// Разрешения считаются только владельцем механизма.
Status.xConfirmAllowed := xRecovery
	AND Input.xPowered
	AND (uiCandidate <> UINT#0)
	AND (Error.dwErrorActive = DWORD#0);
Status.xStartAllowed := Status.xConfirmAllowed
	AND xRobotMagazineReady
	AND xPointsConfigured;
// Общая технологическая готовность не зависит от heartbeat HMI.
xEnableBaseAllowed := xBase
	AND xIdle
	AND Status.xConfirmed
	AND xRobotMagazineReady
	AND xPointsConfigured
	AND (uiCandidate = Status.uiRobotPallet)
	AND Input.xPowered
	AND (Error.dwErrorActive = DWORD#0);
Status.xEnableAllowed := xEnableBaseAllowed AND xConnection;
// Обмен не требует глобальной остановки робота: проверяется только отсутствие
// текущей или уже выданной операции именно с этим магазином.
Status.xSwapAllowed := xBase
	AND xConnection
	AND xIdle
	AND Input.xStandstill
	AND Input.xPowered
	AND (Error.dwErrorActive = DWORD#0)
	AND Status.xConfirmed
	AND (uiCandidate = Status.uiRobotPallet)
	AND NOT Status.xEnabled
	AND NOT xStopRequest
	AND xRobotSwapWindow;
xAutoSwapAllowed := xEnableBaseAllowed
	AND xRobotSwapWindow
	AND Status.xEnabled
	AND xOtherLoaded;
Status.xPowerAllowed := xRecovery
	AND NOT Input.xDriveError
	AND NOT xContradiction;
Status.xDriveResetAllowed := xSelected
	AND xManual
	AND xConnection
	AND Input.xAxisBound
	AND Input.xStandstill
	AND xIdle;
Status.xLowerAllowed := xPneumaticRecovery;
Status.xRaiseAllowed := xRecovery
	AND NOT xContradiction
	AND NOT Status.xHomeRequired;
Status.xSelectAllowed := xRecovery
	AND NOT xContradiction
	AND Input.xLiftDown
	AND NOT Input.xLiftUp
	AND xExchange;
// Наладочные команды замка и фиксатора независимы от подъёма и координаты.
// Это позволяет вернуть герконы в согласованное состояние после остановки.
Status.xLockAllowed := xPneumaticRecovery;
Status.xStopAllowed := xPneumaticRecovery;
Status.xHomeAllowed := xRecovery
	AND Input.xPowered
	AND NOT Input.xDriveError
	AND Input.xLiftDown
	AND NOT Input.xLiftUp
	AND xPairValid
	AND NOT xContradiction;
Status.xMoveAllowed := Status.xHomeAllowed
	AND Input.xHomed
	AND NOT Status.xHomeRequired;
Status.xJogAllowed := Status.xHomeAllowed;
Status.xTeachOperatorAllowed := Status.xMoveAllowed
	AND Input.xLiftDown
	AND NOT Input.xLiftUp;
Status.xTeachWorkAllowed := Status.xTeachOperatorAllowed
	AND ((uiSelected = UINT#1) OR (uiSelected = UINT#2));
Status.xResetAllowed := xRecovery
	AND (Error.dwErrorActive <> DWORD#0)
	AND NOT xContradiction
	AND NOT Input.xDriveError
	AND NOT Status.xHomeRequired
	AND xPairValid
	AND (Input.xLiftDown XOR Input.xLiftUp);
Status.xConfigAllowed := xSelected
	AND xManual
	AND xIdle
	AND NOT Status.xEnabled
	AND (Input.xStandstill OR NOT Input.xAxisBound)
	AND NOT Input.xPowered
	AND NOT xRobotOperation;

// Командный интерфейс FB не зависит от транспортных номеров HMI 1..19.
xCommandPresent := Command.xEnable
	OR Command.xConfirm
	OR Command.xStart
	OR Command.xRejectStart
	OR Command.xDisable
	OR Command.xSwap
	OR Command.xPowerOn
	OR Command.xPowerOff
	OR Command.xDriveReset
	OR Command.xHome
	OR Command.xLower
	OR Command.xRaise
	OR Command.xSelectPallet
	OR Command.xLockIn
	OR Command.xLockOut
	OR Command.xStopIn
	OR Command.xStopOut
	OR Command.xMoveToExchange
	OR Command.xMoveToWork
	OR Command.xStop
	OR Command.xReset
	OR Command.xJogPositive
	OR Command.xJogNegative
	OR Command.xJogRelease
	OR Command.xTeachOperator
	OR Command.xTeachWork;
xAccepted := NOT xCommandPresent;

IF Command.xStart THEN
	IF Status.xStartAllowed
		AND (Command.udiRevision = Status.udiRevision)
		AND (Command.uiPallet = uiCandidate) THEN
		Status.uiRobotPallet := uiCandidate;
		uiConfirmedCandidate := uiCandidate;
		Status.xConfirmed := TRUE;
		Status.xEnabled := TRUE;
		Status.rP1 := 0.0;
		Status.rP2 := 0.0;
		IF uiCandidate = UINT#1 THEN
			Status.rP1 := 1.0;
		ELSE
			Status.rP2 := 1.0;
		END_IF;
		xAccepted := TRUE;
	END_IF;
ELSIF Command.xRejectStart THEN
	Diag.stWarning.uiCode := WRN_START_REJECTED_BY_OPERATOR;
	Diag.stWarning.udiSequence := Diag.stWarning.udiSequence + UDINT#1;
	IF Diag.stWarning.udiSequence = UDINT#0 THEN
		Diag.stWarning.udiSequence := UDINT#1;
	END_IF;
	xAccepted := TRUE;
ELSIF Command.xEnable THEN
	IF Status.xEnableAllowed THEN
		Status.xEnabled := TRUE;
		xAccepted := TRUE;
	END_IF;
ELSIF Command.xConfirm THEN
	IF Status.xConfirmAllowed
		AND (Command.udiRevision = Status.udiRevision)
		AND (Command.uiPallet = uiCandidate) THEN
		Status.uiRobotPallet := uiCandidate;
		uiConfirmedCandidate := uiCandidate;
		Status.xConfirmed := TRUE;
		Status.rP1 := 0.0;
		Status.rP2 := 0.0;
		IF uiCandidate = UINT#1 THEN
			Status.rP1 := 1.0;
		ELSE
			Status.rP2 := 1.0;
		END_IF;
		xAccepted := TRUE;
	END_IF;
ELSIF Command.xDisable THEN
	Status.xEnabled := FALSE;
	xAccepted := TRUE;
ELSIF Command.xSwap THEN
	IF Status.xSwapAllowed THEN
		xExchangeStartedManual := xManual;
		Diag.eState := E_TWO_PALLET_STATE.AUTO_LOWER;
		xAccepted := TRUE;
	END_IF;
ELSIF Command.xPowerOn THEN
	IF Status.xPowerAllowed THEN
		Output.xPowerOn := TRUE;
		xAccepted := TRUE;
	END_IF;
ELSIF Command.xPowerOff THEN
	IF Status.xDriveResetAllowed THEN
		Output.xPowerOff := TRUE;
		Status.xConfirmed := FALSE;
		Status.xEnabled := FALSE;
		xAccepted := TRUE;
	END_IF;
ELSIF Command.xDriveReset THEN
	IF Status.xDriveResetAllowed AND Input.xDriveError THEN
		Output.xDriveReset := TRUE;
		Status.xConfirmed := FALSE;
		Status.xEnabled := FALSE;
		Status.xHomeRequired := TRUE;
		xAccepted := TRUE;
	END_IF;
ELSIF Command.xHome THEN
	IF Status.xHomeAllowed THEN
		Diag.eState := E_TWO_PALLET_STATE.MANUAL_HOME;
		xAccepted := TRUE;
	END_IF;
ELSIF Command.xLower THEN
	IF Status.xLowerAllowed THEN
		Diag.eState := E_TWO_PALLET_STATE.MANUAL_LOWER;
		xAccepted := TRUE;
	END_IF;
ELSIF Command.xRaise THEN
	IF Status.xRaiseAllowed THEN
		Diag.eState := E_TWO_PALLET_STATE.MANUAL_RAISE;
		xAccepted := TRUE;
	END_IF;
ELSIF Command.xSelectPallet THEN
	IF Status.xSelectAllowed
		AND ((Command.uiPallet = UINT#1) OR (Command.uiPallet = UINT#2)) THEN
		uiTo := Command.uiPallet;
		Diag.eState := E_TWO_PALLET_STATE.MANUAL_SELECT_PALLET;
		xAccepted := TRUE;
	END_IF;
ELSIF Command.xLockIn OR Command.xLockOut THEN
	IF Status.xLockAllowed THEN
		xManualLockOutTarget := Command.xLockOut;
		Diag.eState := E_TWO_PALLET_STATE.MANUAL_LOCK;
		xAccepted := TRUE;
	END_IF;
ELSIF Command.xStopIn OR Command.xStopOut THEN
	IF Status.xStopAllowed THEN
		xManualStopOutTarget := Command.xStopOut;
		Diag.eState := E_TWO_PALLET_STATE.MANUAL_STOP;
		xAccepted := TRUE;
	END_IF;
ELSIF Command.xMoveToExchange OR Command.xMoveToWork THEN
	IF Status.xMoveAllowed THEN
		lrTarget := Config.lrExchange;
		IF Command.xMoveToWork THEN
			lrTarget := lrWork;
		END_IF;
		Diag.eState := E_TWO_PALLET_STATE.MANUAL_MOVE;
		xAccepted := TRUE;
	END_IF;
ELSIF Command.xStop THEN
	Status.xEnabled := FALSE;
	// Stop неподвижного механизма не является ручным вмешательством.
	IF (Diag.eState <> E_TWO_PALLET_STATE.IDLE) OR (Input.xPowered AND NOT Input.xStandstill) THEN
		Output.xStop := TRUE;
		Status.xConfirmed := FALSE;
		Error.dwErrorActive := Error.dwErrorActive OR ERR_SEQUENCE_INTERRUPTED;
	END_IF;
	Diag.eState := E_TWO_PALLET_STATE.IDLE;
	uiJogDirection := UINT#0;
	xAccepted := TRUE;
ELSIF Command.xReset THEN
	IF Status.xResetAllowed THEN
		Error.dwErrorLast := Error.dwErrorActive;
		Error.dwErrorActive := DWORD#0;
		Status.xConfirmed := FALSE;
		Status.xEnabled := FALSE;
		xAccepted := TRUE;
	END_IF;
ELSIF Command.xJogPositive OR Command.xJogNegative THEN
	IF Status.xJogAllowed
		OR ((Diag.eState = E_TWO_PALLET_STATE.MANUAL_JOG)
			AND xBase
			AND xManual
			AND xConnection) THEN
		Diag.eState := E_TWO_PALLET_STATE.MANUAL_JOG;
		IF Command.xJogPositive THEN
			uiJogDirection := JOG_POSITIVE;
		ELSE
			uiJogDirection := JOG_NEGATIVE;
		END_IF;
		xAccepted := TRUE;
	END_IF;
ELSIF Command.xJogRelease THEN
	uiJogDirection := UINT#0;
	IF Diag.eState = E_TWO_PALLET_STATE.MANUAL_JOG THEN
		Diag.eState := E_TWO_PALLET_STATE.IDLE;
		Output.xStop := TRUE;
	END_IF;
	xAccepted := TRUE;
ELSIF Command.xTeachOperator THEN
	IF Status.xTeachOperatorAllowed THEN
		Output.xTeachOperator := TRUE;
		xAccepted := TRUE;
	END_IF;
ELSIF Command.xTeachWork THEN
	IF Status.xTeachWorkAllowed THEN
		Output.xTeachWork := TRUE;
		xAccepted := TRUE;
	END_IF;
END_IF;

IF xCommandPresent AND NOT xAccepted THEN
	IF (Command.xEnable OR Command.xStart) AND NOT xPointsConfigured THEN
		Diag.stWarning.uiCode := WRN_ENABLE_POINTS;
	ELSE
		Diag.stWarning.uiCode := WRN_COMMAND_REJECTED;
	END_IF;
	Diag.stWarning.udiSequence := Diag.stWarning.udiSequence + UDINT#1;
	IF Diag.stWarning.udiSequence = UDINT#0 THEN
		Diag.stWarning.udiSequence := UDINT#1;
	END_IF;
END_IF;

IF xExternalCommandRejected THEN
	Diag.stWarning.uiCode := WRN_COMMAND_REJECTED;
	Diag.stWarning.udiSequence := Diag.stWarning.udiSequence + UDINT#1;
	IF Diag.stWarning.udiSequence = UDINT#0 THEN
		Diag.stWarning.udiSequence := UDINT#1;
	END_IF;
END_IF;

Status.xCommandAccepted := xAccepted;

IF xAutoSwap
	AND xAutoSwapAllowed
	AND NOT Output.xStop
	AND NOT xCommandPresent THEN
	xExchangeStartedManual := FALSE;
	Diag.eState := E_TWO_PALLET_STATE.AUTO_LOWER;
END_IF;

// Стоп ячейки имеет приоритет над командой, принятой в том же скане.
// В IDLE при остановленной оси сохраняем включение и подтверждение.
// Собственные Command.xStop / Command.xDisable отдельно отключают магазин.
IF xStopRequest THEN
	IF (Diag.eState <> E_TWO_PALLET_STATE.IDLE) OR (Input.xPowered AND NOT Input.xStandstill) THEN
		Error.dwErrorActive := Error.dwErrorActive OR ERR_SEQUENCE_INTERRUPTED;
		Output.xStop := TRUE;
		Status.xConfirmed := FALSE;
		Status.xEnabled := FALSE;
	END_IF;
	Diag.eState := E_TWO_PALLET_STATE.IDLE;
END_IF;

// Команда могла сменить состояние в этом же скане — обновляем классификацию
// до обработки входа в шаг и запуска таймеров.
xAutomaticState := (Diag.eState = E_TWO_PALLET_STATE.AUTO_LOWER)
	OR (Diag.eState = E_TWO_PALLET_STATE.AUTO_MOVE_TO_EXCHANGE)
	OR (Diag.eState = E_TWO_PALLET_STATE.AUTO_SELECT_PALLET)
	OR (Diag.eState = E_TWO_PALLET_STATE.AUTO_MOVE_TO_WORK)
	OR (Diag.eState = E_TWO_PALLET_STATE.AUTO_RAISE);
xManualState := (Diag.eState = E_TWO_PALLET_STATE.MANUAL_LOWER)
	OR (Diag.eState = E_TWO_PALLET_STATE.MANUAL_RAISE)
	OR (Diag.eState = E_TWO_PALLET_STATE.MANUAL_SELECT_PALLET)
	OR (Diag.eState = E_TWO_PALLET_STATE.MANUAL_MOVE)
	OR (Diag.eState = E_TWO_PALLET_STATE.MANUAL_HOME)
	OR (Diag.eState = E_TWO_PALLET_STATE.MANUAL_JOG)
	OR (Diag.eState = E_TWO_PALLET_STATE.MANUAL_LOCK)
	OR (Diag.eState = E_TWO_PALLET_STATE.MANUAL_STOP);
xManualPneumaticState := (Diag.eState = E_TWO_PALLET_STATE.MANUAL_LOWER)
	OR (Diag.eState = E_TWO_PALLET_STATE.MANUAL_LOCK)
	OR (Diag.eState = E_TWO_PALLET_STATE.MANUAL_STOP);

IF (Diag.eState = E_TWO_PALLET_STATE.AUTO_LOWER)
	AND (ePreviousState <> E_TWO_PALLET_STATE.AUTO_LOWER) THEN
	uiFrom := Status.uiRobotPallet;
	uiTo := UINT#3 - uiFrom;
END_IF;

xStateEntry := Diag.eState <> ePreviousState;
IF xManualState AND xStateEntry THEN
	Status.xConfirmed := FALSE;
	Status.xEnabled := FALSE;
	Status.udiRevision := Status.udiRevision + UDINT#1;
	IF Status.udiRevision = UDINT#0 THEN
		Status.udiRevision := UDINT#1;
	END_IF;
END_IF;

IF xStateEntry THEN
	xSeenMotion := FALSE;
	xSeenDone := FALSE;
	IF (Diag.eState = E_TWO_PALLET_STATE.MANUAL_MOVE)
		OR (Diag.eState = E_TWO_PALLET_STATE.MANUAL_HOME)
		OR (Diag.eState = E_TWO_PALLET_STATE.MANUAL_JOG) THEN
		uiManualSelected := uiSelected;
	END_IF;
ELSIF Input.xMotionDone THEN
	xSeenDone := TRUE;
END_IF;

IF NOT Input.xStandstill THEN
	xSeenMotion := TRUE;
END_IF;

tStateLimit := Config.tCylinder;
IF (Diag.eState = E_TWO_PALLET_STATE.AUTO_MOVE_TO_EXCHANGE)
	OR (Diag.eState = E_TWO_PALLET_STATE.AUTO_MOVE_TO_WORK)
	OR (Diag.eState = E_TWO_PALLET_STATE.MANUAL_MOVE) THEN
	tStateLimit := Config.tMove;
END_IF;
IF Diag.eState = E_TWO_PALLET_STATE.MANUAL_HOME THEN
	tStateLimit := Config.tHome;
END_IF;

tonState(
	IN := NOT xIdle
		AND (Diag.eState <> E_TWO_PALLET_STATE.MANUAL_JOG)
		AND NOT xStateEntry,
	PT := tStateLimit);
tonCoil(
	IN := NOT xIdle AND NOT xStateEntry,
	PT := Config.tPulse);
tonJogLease(
	IN := (Diag.eState = E_TWO_PALLET_STATE.MANUAL_JOG)
		AND NOT (Command.xJogPositive OR Command.xJogNegative),
	PT := T#350MS);
ePreviousState := Diag.eState;

// Автомат обмена и ручного восстановления.
uiTargetSignals := Config.uiP1Signals;
IF uiTo = UINT#2 THEN uiTargetSignals := Config.uiP2Signals; END_IF;
CASE Diag.eState OF
	E_TWO_PALLET_STATE.AUTO_LOWER,
	E_TWO_PALLET_STATE.MANUAL_LOWER:
		xLiftDownCommand := TRUE;
		IF Input.xLiftDown AND NOT Input.xLiftUp THEN
			IF Diag.eState = E_TWO_PALLET_STATE.AUTO_LOWER THEN
				Diag.eState := E_TWO_PALLET_STATE.AUTO_MOVE_TO_EXCHANGE;
				lrTarget := Config.lrExchange;
			ELSE
				Diag.eState := E_TWO_PALLET_STATE.IDLE;
			END_IF;
		END_IF;

	E_TWO_PALLET_STATE.AUTO_MOVE_TO_EXCHANGE,
	E_TWO_PALLET_STATE.AUTO_MOVE_TO_WORK,
	E_TWO_PALLET_STATE.MANUAL_MOVE:
		IF Diag.eState = E_TWO_PALLET_STATE.AUTO_MOVE_TO_WORK THEN
			lrTarget := Config.lrWorkP1;
			IF uiTo = UINT#2 THEN
				lrTarget := Config.lrWorkP2;
			END_IF;
		END_IF;

		IF NOT Input.xLiftDown
			OR Input.xLiftUp
			OR NOT xPairValid
			OR Status.xHomeRequired
			OR ((Diag.eState = E_TWO_PALLET_STATE.AUTO_MOVE_TO_EXCHANGE) AND (uiSelected <> uiFrom))
			OR ((Diag.eState = E_TWO_PALLET_STATE.AUTO_MOVE_TO_WORK) AND (uiSelected <> uiTo))
			OR ((Diag.eState = E_TWO_PALLET_STATE.MANUAL_MOVE) AND (uiSelected <> uiManualSelected))
			OR (Input.xLimitPositive AND (lrTarget > Input.lrPosition + Config.lrTolerance))
			OR (Input.xLimitNegative AND (lrTarget < Input.lrPosition - Config.lrTolerance)) THEN
			Error.dwErrorActive := Error.dwErrorActive OR ERR_LOGIC;
			Diag.eState := E_TWO_PALLET_STATE.IDLE;
			Output.xStop := TRUE;
		ELSE
			Output.lrTarget := lrTarget;
			Output.xMove := xStateEntry;
			IF Input.xStandstill
				AND (ABS(Input.lrPosition - lrTarget) <= Config.lrTolerance)
				AND ((xSeenMotion OR xSeenDone) OR xStateEntry) THEN
				Output.xMove := FALSE;
				IF Diag.eState = E_TWO_PALLET_STATE.AUTO_MOVE_TO_EXCHANGE THEN
					Diag.eState := E_TWO_PALLET_STATE.AUTO_SELECT_PALLET;
				ELSIF Diag.eState = E_TWO_PALLET_STATE.AUTO_MOVE_TO_WORK THEN
					Diag.eState := E_TWO_PALLET_STATE.AUTO_RAISE;
				ELSE
					Diag.eState := E_TWO_PALLET_STATE.IDLE;
				END_IF;
			END_IF;
		END_IF;

	E_TWO_PALLET_STATE.AUTO_SELECT_PALLET,
	E_TWO_PALLET_STATE.MANUAL_SELECT_PALLET:
		IF NOT xExchange OR NOT Input.xLiftDown OR Input.xLiftUp THEN
			Error.dwErrorActive := Error.dwErrorActive OR ERR_LOGIC;
			Diag.eState := E_TWO_PALLET_STATE.IDLE;
			Output.xStop := TRUE;
		ELSE
			xSelectCommand := TRUE;
		END_IF;
		IF (uiSelected = uiTo) AND xPairValid AND NOT Output.xStop THEN
			IF Diag.eState = E_TWO_PALLET_STATE.AUTO_SELECT_PALLET THEN
				Diag.eState := E_TWO_PALLET_STATE.AUTO_MOVE_TO_WORK;
			ELSE
				Diag.eState := E_TWO_PALLET_STATE.IDLE;
			END_IF;
		END_IF;

	E_TWO_PALLET_STATE.MANUAL_LOCK:
		IF xManualLockOutTarget THEN
			xManualLockCommand := NOT Input.xLockOut OR Input.xLockIn;
			IF Input.xLockOut AND NOT Input.xLockIn THEN Diag.eState := E_TWO_PALLET_STATE.IDLE; END_IF;
		ELSE
			xManualLockCommand := NOT Input.xLockIn OR Input.xLockOut;
			IF Input.xLockIn AND NOT Input.xLockOut THEN Diag.eState := E_TWO_PALLET_STATE.IDLE; END_IF;
		END_IF;

	E_TWO_PALLET_STATE.MANUAL_STOP:
		IF xManualStopOutTarget THEN
			xManualStopCommand := NOT Input.xStopOut OR Input.xStopIn;
			IF Input.xStopOut AND NOT Input.xStopIn THEN Diag.eState := E_TWO_PALLET_STATE.IDLE; END_IF;
		ELSE
			xManualStopCommand := NOT Input.xStopIn OR Input.xStopOut;
			IF Input.xStopIn AND NOT Input.xStopOut THEN Diag.eState := E_TWO_PALLET_STATE.IDLE; END_IF;
		END_IF;

	E_TWO_PALLET_STATE.AUTO_RAISE:
		// Завершение обмена устанавливает подъём по выбранной конфигурации
		// только после фактического останова в рабочей позиции.
		IF NOT xWork
			OR Status.xHomeRequired
			OR (uiSelected <> uiTo) THEN
			Error.dwErrorActive := Error.dwErrorActive OR ERR_LOGIC;
			Diag.eState := E_TWO_PALLET_STATE.IDLE;
			Output.xStop := TRUE;
		ELSE
			xLiftUpCommand := (uiTargetSignals AND UINT#2) <> UINT#0;
			xLiftDownCommand := NOT xLiftUpCommand;
			IF uiSignals = uiTargetSignals THEN
				Status.uiRobotPallet := uiTo;
				uiConfirmedCandidate := uiTo;
				Status.xConfirmed := TRUE;
				Status.xCompleted := TRUE;
				Diag.eState := E_TWO_PALLET_STATE.IDLE;
			END_IF;
		END_IF;

	E_TWO_PALLET_STATE.MANUAL_RAISE:
		// Наладочный подъём не требует HOME-координаты или рабочей позиции.
		IF NOT Input.xStandstill OR NOT xManual OR xContradiction OR Status.xHomeRequired THEN
			Error.dwErrorActive := Error.dwErrorActive OR ERR_LOGIC;
			Diag.eState := E_TWO_PALLET_STATE.IDLE;
			Output.xStop := TRUE;
		ELSE
			xLiftUpCommand := TRUE;
			IF Input.xLiftUp AND NOT Input.xLiftDown THEN
				Diag.eState := E_TWO_PALLET_STATE.IDLE;
			END_IF;
		END_IF;

	E_TWO_PALLET_STATE.MANUAL_HOME:
		Output.xHome := xStateEntry;
		IF xSeenDone
			AND Input.xHomed
			AND Input.xStandstill
			AND NOT xStateEntry THEN
			Status.xHomeRequired := FALSE;
			Diag.eState := E_TWO_PALLET_STATE.IDLE;
		END_IF;

	E_TWO_PALLET_STATE.MANUAL_JOG:
		IF tonJogLease.Q OR NOT xConnection OR (uiJogDirection = UINT#0) THEN
			Diag.eState := E_TWO_PALLET_STATE.IDLE;
			Output.xStop := TRUE;
		ELSE
			Output.xJogPositive := (uiJogDirection = JOG_POSITIVE) AND NOT Input.xLimitPositive;
			Output.xJogNegative := (uiJogDirection = JOG_NEGATIVE) AND NOT Input.xLimitNegative;
		END_IF;

	E_TWO_PALLET_STATE.IDLE:
		uiJogDirection := UINT#0;

ELSE
	Error.dwErrorActive := Error.dwErrorActive OR ERR_LOGIC;
	Diag.eState := E_TWO_PALLET_STATE.IDLE;
	Output.xStop := TRUE;
END_CASE;
IF Diag.eState = E_TWO_PALLET_STATE.IDLE THEN xExchangeStartedManual := FALSE; END_IF;

// Низ П2 и выбранное зацепление контролируются всё время Home/JOG.
IF ((Diag.eState = E_TWO_PALLET_STATE.MANUAL_HOME)
	OR (Diag.eState = E_TWO_PALLET_STATE.MANUAL_JOG))
	AND (NOT Input.xLiftDown
		OR Input.xLiftUp
		OR NOT xPairValid
		OR (uiSelected <> uiManualSelected)
		OR xContradiction
		OR Input.xDriveError
		OR NOT Input.xPowered) THEN
	Error.dwErrorActive := Error.dwErrorActive OR ERR_LOGIC;
	Diag.eState := E_TWO_PALLET_STATE.IDLE;
	Output.xStop := TRUE;
END_IF;

IF tonState.Q THEN
	IF (ePreviousState = E_TWO_PALLET_STATE.AUTO_MOVE_TO_EXCHANGE)
		OR (ePreviousState = E_TWO_PALLET_STATE.AUTO_MOVE_TO_WORK)
		OR (ePreviousState = E_TWO_PALLET_STATE.MANUAL_MOVE)
		OR (ePreviousState = E_TWO_PALLET_STATE.MANUAL_HOME) THEN
		Error.dwErrorActive := Error.dwErrorActive OR ERR_MOTION_TIMEOUT;
		Status.xHomeRequired := TRUE;
	ELSE
		Error.dwErrorActive := Error.dwErrorActive OR ERR_CYLINDER_TIMEOUT;
	END_IF;
	Diag.eState := E_TWO_PALLET_STATE.IDLE;
	Output.xStop := TRUE;
END_IF;

IF (((NOT xBase) AND NOT (xManualPneumaticState AND xPneumaticBase))
	OR ((NOT xConnection) AND xManualState AND NOT xManualPneumaticState))
	AND (ePreviousState <> E_TWO_PALLET_STATE.IDLE)
	OR Output.xStop THEN
	Output.xMove := FALSE;
	Output.xHome := FALSE;
	Output.xJogPositive := FALSE;
	Output.xJogNegative := FALSE;
	xLiftUpCommand := FALSE;
	xLiftDownCommand := FALSE;
	xSelectCommand := FALSE;
	xManualLockCommand := FALSE;
	xManualStopCommand := FALSE;
END_IF;

// Автоматический обмен переключает пару совместно; ручное восстановление — каждый цилиндр отдельно.
xLockOutTarget := (uiTargetSignals AND UINT#8) <> UINT#0;
xStopOutTarget := (uiTargetSignals AND UINT#32) <> UINT#0;
Output.xLiftUp := xBase AND xLiftUpCommand AND NOT tonCoil.Q;
Output.xLiftDown := (xBase OR xPneumaticBase) AND xLiftDownCommand AND NOT tonCoil.Q;
Output.xLockOut := (xBase AND xSelectCommand AND xLockOutTarget
	OR xPneumaticBase AND xManualLockCommand AND xManualLockOutTarget) AND NOT tonCoil.Q;
Output.xLockIn := (xBase AND xSelectCommand AND NOT xLockOutTarget
	OR xPneumaticBase AND xManualLockCommand AND NOT xManualLockOutTarget) AND NOT tonCoil.Q;
Output.xStopOut := (xBase AND xSelectCommand AND xStopOutTarget
	OR xPneumaticBase AND xManualStopCommand AND xManualStopOutTarget) AND NOT tonCoil.Q;
Output.xStopIn := (xBase AND xSelectCommand AND NOT xStopOutTarget
	OR xPneumaticBase AND xManualStopCommand AND NOT xManualStopOutTarget) AND NOT tonCoil.Q;

// Поза для 3D — оценка по координате каретки и подтверждённому зацеплению.
IF xPairValid AND Input.xHomed THEN
	lrSpan := lrWork - Config.lrExchange;
	IF ABS(lrSpan) > Config.lrTolerance THEN
		rTravel := LREAL_TO_REAL(
			LIMIT(0.0, (Input.lrPosition - Config.lrExchange) / lrSpan, 1.0));
		IF uiSelected = UINT#1 THEN
			Status.rP1 := rTravel;
		ELSE
			Status.rP2 := rTravel;
		END_IF;
	END_IF;
END_IF;

IF Input.xLiftUp AND NOT Input.xLiftDown THEN
	Status.rLift := 1.0;
ELSIF Input.xLiftDown AND NOT Input.xLiftUp THEN
	Status.rLift := 0.0;
END_IF;

// Диагностика и совместимый публичный Status формируются в одном месте.
IF (Error.dwErrorActive <> dwPreviousError)
	AND (Error.dwErrorActive <> DWORD#0) THEN
	Diag.eFaultState := ePreviousState;
END_IF;
dwPreviousError := Error.dwErrorActive;

IF Error.dwErrorActive <> DWORD#0 THEN
	Error.dwErrorLast := Error.dwErrorActive;
	Status.xConfirmed := FALSE;
	Status.xEnabled := FALSE;
END_IF;
Error.dwAlarmActive := Error.dwErrorActive;
Error.stErrorActive := UpdateErrorView(dwError := Error.dwErrorActive);
Error.stErrorLast := UpdateErrorView(dwError := Error.dwErrorLast);

Status.uiStep := TO_UINT(Diag.eState);
Status.uiFaultStep := TO_UINT(Diag.eFaultState);
Status.uiReason := Diag.uiReason;
Status.dwError := Error.dwErrorActive;
Status.stWarning := Diag.stWarning;
Status.xBusy := Diag.eState <> E_TWO_PALLET_STATE.IDLE;
Status.xError := Error.dwErrorActive <> DWORD#0;

// Команда или автомат могли занять механизм после первоначального расчёта
// разрешений. Не публикуем устаревшее разрешение ещё на один скан.
IF Status.xBusy THEN
	Status.xConfirmAllowed := FALSE;
	Status.xStartAllowed := FALSE;
	Status.xEnableAllowed := FALSE;
	Status.xSwapAllowed := FALSE;
	Status.xPowerAllowed := FALSE;
	Status.xDriveResetAllowed := FALSE;
	Status.xHomeAllowed := FALSE;
	Status.xLowerAllowed := FALSE;
	Status.xRaiseAllowed := FALSE;
	Status.xSelectAllowed := FALSE;
	Status.xLockAllowed := FALSE;
	Status.xStopAllowed := FALSE;
	Status.xMoveAllowed := FALSE;
	Status.xJogAllowed := FALSE;
	Status.xTeachOperatorAllowed := FALSE;
	Status.xTeachWorkAllowed := FALSE;
	Status.xResetAllowed := FALSE;
	Status.xConfigAllowed := FALSE;
END_IF;

// Инвентарь операторской палеты редактируется всегда, независимо от режима,
// движения, подтверждения, питания и ошибок механизма. Роботная палета — только
// при выключенном магазине после освобождения текущей/выданной операции с ним.
// Считаем после команд и обмена, чтобы роль палеты была актуальна в этом скане.
Status.xEdit1Allowed := xSelected
	AND ((Status.uiRobotPallet <> UINT#1) OR (NOT Status.xEnabled AND xActivePalletEditAllowed));
Status.xEdit2Allowed := xSelected
	AND ((Status.uiRobotPallet <> UINT#2) OR (NOT Status.xEnabled AND xActivePalletEditAllowed));
Status.xEditAllowed := Status.xEdit1Allowed OR Status.xEdit2Allowed;
Status.xLoadAllowed := Status.xConfirmed AND NOT Status.xBusy AND NOT xOtherLoaded
	AND (((Status.uiRobotPallet = UINT#1) AND Status.xEdit2Allowed)
		OR ((Status.uiRobotPallet = UINT#2) AND Status.xEdit1Allowed));

Status.xReady := xSelected
	AND Status.xEnabled
	AND Status.xConfirmed
	AND NOT Status.xBusy
	AND NOT Status.xError
	AND xWork
	AND (uiCandidate = Status.uiRobotPallet)
	AND Input.xPowered
	AND xRobotGeometryReady
	AND xRobotMagazineReady
	AND xSafe;

IF NOT xSelected THEN
	Status.xEnabled := FALSE;
	Status.xConfirmed := FALSE;
END_IF;

METHOD IsSignalConfigurationValid : BOOL
VAR_INPUT
	uiP1Signals : UINT;
	uiP2Signals : UINT;
END_VAR
// Рабочее положение каждого цилиндра подтверждает ровно один геркон.
// Зацепление должно различать палеты и при опущенной П2 во время обмена.
IsSignalConfigurationValid := (uiP1Signals <= UINT#63)
	AND (uiP2Signals <= UINT#63)
	AND (((uiP1Signals AND UINT#3) = UINT#1) OR ((uiP1Signals AND UINT#3) = UINT#2))
	AND (((uiP2Signals AND UINT#3) = UINT#1) OR ((uiP2Signals AND UINT#3) = UINT#2))
	AND (((uiP1Signals AND UINT#12) = UINT#4) OR ((uiP1Signals AND UINT#12) = UINT#8))
	AND (((uiP2Signals AND UINT#12) = UINT#4) OR ((uiP2Signals AND UINT#12) = UINT#8))
	AND (((uiP1Signals AND UINT#48) = UINT#16) OR ((uiP1Signals AND UINT#48) = UINT#32))
	AND (((uiP2Signals AND UINT#48) = UINT#16) OR ((uiP2Signals AND UINT#48) = UINT#32))
	AND ((uiP1Signals AND UINT#60) <> (uiP2Signals AND UINT#60));
END_METHOD

METHOD UpdateErrorView : ST_TWO_PALLET_ERROR
VAR_INPUT
	dwError : DWORD;
END_VAR
VAR
	stError : ST_TWO_PALLET_ERROR;
END_VAR
stError.DRIVE_ERROR := (dwError AND ERR_DRIVE) <> DWORD#0;
stError.SENSOR_CONTRADICTION := (dwError AND ERR_SENSOR_CONTRADICTION) <> DWORD#0;
stError.CYLINDER_TIMEOUT := (dwError AND ERR_CYLINDER_TIMEOUT) <> DWORD#0;
stError.MOTION_TIMEOUT := (dwError AND ERR_MOTION_TIMEOUT) <> DWORD#0;
stError.LOGIC_ERROR := (dwError AND ERR_LOGIC) <> DWORD#0;
stError.SEQUENCE_INTERRUPTED := (dwError AND ERR_SEQUENCE_INTERRUPTED) <> DWORD#0;

UpdateErrorView := stError;
END_METHOD

END_FUNCTION_BLOCK

// Device/Application/FB/FB_TWO_PALLET_SIMULATION
FUNCTION_BLOCK FB_TWO_PALLET_SIMULATION
VAR_INPUT
	xEnable : BOOL; // Только тестовая среда SIMULATION
	uiP1Signals : UINT;
	Command : ST_TWO_PALLET_OUTPUT;
END_VAR
VAR_OUTPUT
	xLiftDown : BOOL;
	xLiftUp : BOOL;
	xLockIn : BOOL;
	xLockOut : BOOL;
	xStopIn : BOOL;
	xStopOut : BOOL;
END_VAR
VAR
	xInitialized : BOOL;
	xLiftTargetUp : BOOL;
	xLockTargetOut : BOOL;
	xStopTargetOut : BOOL;
	tonLift : TON;
	tonLock : TON;
	tonStop : TON;
END_VAR

IF NOT xEnable THEN
	xInitialized := FALSE;
	xLiftDown := FALSE;
	xLiftUp := FALSE;
	xLockIn := FALSE;
	xLockOut := FALSE;
	xStopIn := FALSE;
	xStopOut := FALSE;
	tonLift(IN := FALSE, PT := T#300MS);
	tonLock(IN := FALSE, PT := T#300MS);
	tonStop(IN := FALSE, PT := T#300MS);
ELSE
	IF NOT xInitialized THEN
		// Виртуальная начальная поза: П2 внизу, замок держит П1,
		// фиксатор держит противоположную палету.
		xLiftTargetUp := FALSE;
		xLockTargetOut := (uiP1Signals AND UINT#8) <> UINT#0;
		xStopTargetOut := (uiP1Signals AND UINT#32) <> UINT#0;
		xLiftDown := TRUE;
		xLiftUp := FALSE;
		xLockOut := xLockTargetOut;
		xLockIn := NOT xLockTargetOut;
		xStopOut := xStopTargetOut;
		xStopIn := NOT xStopTargetOut;
		xInitialized := TRUE;
	END_IF;

	// Бистабильный 5/2 сохраняет положение после снятия обеих катушек.
	IF Command.xLiftUp AND NOT Command.xLiftDown THEN
		xLiftTargetUp := TRUE;
	ELSIF Command.xLiftDown AND NOT Command.xLiftUp THEN
		xLiftTargetUp := FALSE;
	END_IF;
	IF Command.xLockOut AND NOT Command.xLockIn THEN
		xLockTargetOut := TRUE;
	ELSIF Command.xLockIn AND NOT Command.xLockOut THEN
		xLockTargetOut := FALSE;
	END_IF;
	IF Command.xStopOut AND NOT Command.xStopIn THEN
		xStopTargetOut := TRUE;
	ELSIF Command.xStopIn AND NOT Command.xStopOut THEN
		xStopTargetOut := FALSE;
	END_IF;

	tonLift(IN := xLiftTargetUp <> xLiftUp, PT := T#300MS);
	tonLock(IN := xLockTargetOut <> xLockOut, PT := T#300MS);
	tonStop(IN := xStopTargetOut <> xStopOut, PT := T#300MS);
	IF tonLift.Q THEN
		xLiftUp := xLiftTargetUp;
		xLiftDown := NOT xLiftTargetUp;
	END_IF;
	IF tonLock.Q THEN
		xLockOut := xLockTargetOut;
		xLockIn := NOT xLockTargetOut;
	END_IF;
	IF tonStop.Q THEN
		xStopOut := xStopTargetOut;
		xStopIn := NOT xStopTargetOut;
	END_IF;
END_IF;

END_FUNCTION_BLOCK

// Device/Application/FB/FB_MULTI_TYPE/FB_MULTI_TYPE_CONFIG_MANAGER
FUNCTION_BLOCK FB_MULTI_TYPE_CONFIG_MANAGER
VAR_INPUT
	xTestInitialize  : BOOL; // Атомарная загрузка конфигурации из тестового буфера
	stTestScenario   : ST_TEST_SCENARIO_BUFFER;
	Command          : ST_MULTI_TYPE_COMMAND; // Запросы конфигурации от HMI
	xCellRunning     : BOOL; // Автоматический цикл выполняется
	xMotionBusy      : BOOL; // Оси ещё движутся
	stRobotStatus    : ST_ROBOT_STATUS; // Состояние робота
	astMagazineStatus : ARRAY [1..GVL_CELL_SETTINGS.MagazineCount] OF ST_MAGAZINE_STATUS; // Оба магазина
	astMachineStatus : ARRAY [1..3] OF ST_MACHINE_PUBLIC; // Состояния станков
	uiRows           : UINT; // Строки активной матрицы
	uiColumns        : UINT; // Столбцы активной матрицы
END_VAR
VAR_OUTPUT
	Config : ST_MULTI_TYPE_CONFIG; // Фактически принятая конфигурация
	Status : ST_MULTI_TYPE_CONFIG_STATUS; // Разрешения и диагностика
END_VAR
VAR
	xInitialized        : BOOL; // Начальные безопасные значения заданы
	xAllMachinesSafe    : BOOL; // Станки не обслуживаются и не обрабатывают
	xAllMachinesDisabled: BOOL; // Все станки выключены
	xAllMagazinesEditable : BOOL; // Оба магазина выключены и не заняты
	xAllTypesHaveMachines : BOOL; // Каждый тип назначен хотя бы одному станку
	uiMachine           : UINT; // Индекс станка
	uiMagazine          : UINT; // Индекс магазина
	uiSlot              : UINT; // Индекс слота
	uiType              : UINT; // Индекс типа
	auiMachineCount     : ARRAY [1..3] OF UINT; // Количество станков каждого типа
	auiSlotCount        : ARRAY [1..3] OF UINT; // Количество слотов каждого типа
	rtSetTypeCount      : R_TRIG; // Фронт изменения количества типов
	rtSetMachineType    : R_TRIG; // Фронт назначения типа станку
	rtSetSlotType       : R_TRIG; // Фронт назначения типа слоту
	rtAutoDistribute    : R_TRIG; // Фронт автоматического распределения
END_VAR
VAR CONSTANT
	FIRST_MACHINE : UINT := UINT#1;
	LAST_MACHINE  : UINT := UINT#3;
	FIRST_TYPE    : UINT := UINT#1;
	LAST_TYPE     : UINT := UINT#3;
	WRN_TYPE_COUNT_NOT_ALLOWED : UINT := UINT#23;
	WRN_MACHINE_TYPE_REJECTED  : UINT := UINT#24;
	WRN_SLOT_TYPE_REJECTED     : UINT := UINT#25;
	WRN_DISTRIBUTION_REJECTED  : UINT := UINT#26;
END_VAR

IF (uiRows > UINT#0)
AND (uiColumns > UINT#0)
AND ((uiRows * uiColumns) <= SINT_TO_UINT(GVL_CELL_SETTINGS.NumberDetail)) THEN
	Status.uiActiveSlotCount := uiRows * uiColumns;
ELSE
	Status.uiActiveSlotCount := UINT#0;
END_IF;

IF NOT xInitialized THEN
	Config.uiTypeCount := UINT#1;
	FOR uiMachine := FIRST_MACHINE TO LAST_MACHINE DO
		Config.auiMachineType[uiMachine] := UINT#1;
	END_FOR;
	FOR uiSlot := UINT#1 TO SINT_TO_UINT(GVL_CELL_SETTINGS.NumberDetail) DO
		IF uiSlot <= Status.uiActiveSlotCount THEN
			Config.auiSlotType[uiSlot] := UINT#1;
		ELSE
			Config.auiSlotType[uiSlot] := UINT#0;
		END_IF;
	END_FOR;
	xInitialized := TRUE;
END_IF;

xAllMachinesSafe := TRUE;
xAllMachinesDisabled := TRUE;
FOR uiMachine := FIRST_MACHINE TO LAST_MACHINE DO
	IF astMachineStatus[uiMachine].xBusy
	OR astMachineStatus[uiMachine].xProcessing THEN
		xAllMachinesSafe := FALSE;
	END_IF;
	IF astMachineStatus[uiMachine].xEnabled
	OR astMachineStatus[uiMachine].xDisablePending THEN
		xAllMachinesDisabled := FALSE;
	END_IF;
END_FOR;

xAllMagazinesEditable := TRUE;
FOR uiMagazine := UINT#1 TO INT_TO_UINT(GVL_CELL_SETTINGS.MagazineCount) DO
	IF astMagazineStatus[uiMagazine].xEnabled
	OR astMagazineStatus[uiMagazine].xBusy
	OR astMagazineStatus[uiMagazine].xDisablePending THEN
		xAllMagazinesEditable := FALSE;
	END_IF;
END_FOR;

Status.xMagazineConfigAllowed := NOT xCellRunning
	AND NOT xMotionBusy
	AND NOT stRobotStatus.xBusy
	AND NOT stRobotStatus.xBlankAvailable
	AND NOT stRobotStatus.xDetailAvailable
	AND xAllMagazinesEditable
	AND xAllMachinesSafe;
Status.xTypeCountAllowed := Status.xMagazineConfigAllowed
	AND xAllMachinesDisabled;

FOR uiMachine := FIRST_MACHINE TO LAST_MACHINE DO
	Status.axMachineTypeAllowed[uiMachine] := NOT xCellRunning
		AND NOT xMotionBusy
		AND NOT stRobotStatus.xBusy
		AND NOT stRobotStatus.xBlankAvailable
		AND NOT stRobotStatus.xDetailAvailable
		AND xAllMagazinesEditable
		AND NOT astMachineStatus[uiMachine].xEnabled
		AND NOT astMachineStatus[uiMachine].xDisablePending
		AND NOT astMachineStatus[uiMachine].xBusy
		AND NOT astMachineStatus[uiMachine].xProcessing;
END_FOR;

rtSetTypeCount(CLK := Command.xSetTypeCount);
rtSetMachineType(CLK := Command.xSetMachineType);
rtSetSlotType(CLK := Command.xSetSlotType);
rtAutoDistribute(CLK := Command.xAutoDistribute);

IF rtSetTypeCount.Q THEN
	IF NOT Status.xTypeCountAllowed
	OR (Command.uiRequestedTypeCount < FIRST_TYPE)
	OR (Command.uiRequestedTypeCount > LAST_TYPE) THEN
		RaiseWarning(uiCode := WRN_TYPE_COUNT_NOT_ALLOWED);
	ELSE
		Config.uiTypeCount := Command.uiRequestedTypeCount;
		CASE Config.uiTypeCount OF
			UINT#1:
				Config.auiMachineType[1] := UINT#1;
				Config.auiMachineType[2] := UINT#1;
				Config.auiMachineType[3] := UINT#1;
			UINT#2:
				Config.auiMachineType[1] := UINT#1;
				Config.auiMachineType[2] := UINT#1;
				Config.auiMachineType[3] := UINT#2;
			UINT#3:
				Config.auiMachineType[1] := UINT#1;
				Config.auiMachineType[2] := UINT#2;
				Config.auiMachineType[3] := UINT#3;
		END_CASE;
		ApplyDistribution();
	END_IF;
END_IF;

IF rtSetMachineType.Q THEN
	IF (Command.uiRequestedMachine < FIRST_MACHINE)
	OR (Command.uiRequestedMachine > LAST_MACHINE) THEN
		RaiseWarning(uiCode := WRN_MACHINE_TYPE_REJECTED);
	ELSE
		IF (Command.uiRequestedMachineType < FIRST_TYPE)
		OR (Command.uiRequestedMachineType > Config.uiTypeCount)
		OR NOT Status.axMachineTypeAllowed[Command.uiRequestedMachine] THEN
			RaiseWarning(uiCode := WRN_MACHINE_TYPE_REJECTED);
		ELSE
			Config.auiMachineType[Command.uiRequestedMachine] := Command.uiRequestedMachineType;
		END_IF;
	END_IF;
END_IF;

IF rtSetSlotType.Q THEN
	IF NOT Status.xMagazineConfigAllowed
	OR (Command.uiRequestedSlot < UINT#1)
	OR (Command.uiRequestedSlot > Status.uiActiveSlotCount)
	OR (Command.uiRequestedSlotType < FIRST_TYPE)
	OR (Command.uiRequestedSlotType > Config.uiTypeCount) THEN
		RaiseWarning(uiCode := WRN_SLOT_TYPE_REJECTED);
	ELSE
		Config.auiSlotType[Command.uiRequestedSlot] := Command.uiRequestedSlotType;
	END_IF;
END_IF;

IF rtAutoDistribute.Q THEN
	xAllTypesHaveMachines := TRUE;
	FOR uiType := FIRST_TYPE TO LAST_TYPE DO
		auiMachineCount[uiType] := UINT#0;
	END_FOR;
	FOR uiMachine := FIRST_MACHINE TO LAST_MACHINE DO
		IF (Config.auiMachineType[uiMachine] >= FIRST_TYPE)
		AND (Config.auiMachineType[uiMachine] <= Config.uiTypeCount) THEN
			auiMachineCount[Config.auiMachineType[uiMachine]] :=
				auiMachineCount[Config.auiMachineType[uiMachine]] + UINT#1;
		END_IF;
	END_FOR;
	FOR uiType := FIRST_TYPE TO Config.uiTypeCount DO
		IF auiMachineCount[uiType] = UINT#0 THEN
			xAllTypesHaveMachines := FALSE;
		END_IF;
	END_FOR;

	IF NOT Status.xMagazineConfigAllowed
	OR NOT xAllTypesHaveMachines THEN
		RaiseWarning(uiCode := WRN_DISTRIBUTION_REJECTED);
	ELSE
		ApplyDistribution();
	END_IF;
END_IF;

// Тестовый сценарий проходит общую PLC-валидацию до этого вызова. Запись
// выполняет владелец Config, поэтому значения не теряются на выходной привязке FB.
IF xTestInitialize THEN
	Config.uiTypeCount := stTestScenario.uiTypeCount;
	FOR uiMachine := FIRST_MACHINE TO LAST_MACHINE DO
		Config.auiMachineType[uiMachine] := stTestScenario.auiMachineType[uiMachine];
	END_FOR;
	FOR uiSlot := UINT#1 TO SINT_TO_UINT(GVL_CELL_SETTINGS.NumberDetail) DO
		Config.auiSlotType[uiSlot] := stTestScenario.auiSlotType[uiSlot];
	END_FOR;
END_IF;

FOR uiType := FIRST_TYPE TO LAST_TYPE DO
	auiMachineCount[uiType] := UINT#0;
	auiSlotCount[uiType] := UINT#0;
END_FOR;

Status.xConfigurationValid := (Config.uiTypeCount >= FIRST_TYPE)
	AND (Config.uiTypeCount <= LAST_TYPE)
	AND (Status.uiActiveSlotCount > UINT#0);

FOR uiMachine := FIRST_MACHINE TO LAST_MACHINE DO
	IF (Config.auiMachineType[uiMachine] < FIRST_TYPE)
	OR (Config.auiMachineType[uiMachine] > Config.uiTypeCount) THEN
		Status.xConfigurationValid := FALSE;
	ELSE
		auiMachineCount[Config.auiMachineType[uiMachine]] :=
			auiMachineCount[Config.auiMachineType[uiMachine]] + UINT#1;
	END_IF;
END_FOR;

FOR uiSlot := UINT#1 TO Status.uiActiveSlotCount DO
	IF (Config.auiSlotType[uiSlot] < FIRST_TYPE)
	OR (Config.auiSlotType[uiSlot] > Config.uiTypeCount) THEN
		Status.xConfigurationValid := FALSE;
	ELSE
		auiSlotCount[Config.auiSlotType[uiSlot]] :=
			auiSlotCount[Config.auiSlotType[uiSlot]] + UINT#1;
	END_IF;
END_FOR;

FOR uiType := FIRST_TYPE TO Config.uiTypeCount DO
	IF (auiMachineCount[uiType] = UINT#0)
	OR (auiSlotCount[uiType] = UINT#0) THEN
		Status.xConfigurationValid := FALSE;
	END_IF;
END_FOR;

METHOD PRIVATE ApplyDistribution
VAR
	uiMachine       : UINT; // Индекс станка
	uiType          : UINT; // Индекс типа
	uiSlot          : UINT; // Индекс слота
	uiAssigned      : UINT; // Число уже назначенных слотов
	uiRemaining     : UINT; // Остаток после целочисленного деления
	uiBestType      : UINT; // Тип с наибольшей дробной частью
	uiBestRemainder : UINT; // Наибольшая дробная часть
	auiMachineShare : ARRAY [1..3] OF UINT; // Число станков типа
	auiQuota        : ARRAY [1..3] OF UINT; // Число слотов типа
	auiRemainder    : ARRAY [1..3] OF UINT; // Остаток квоты
	axExtraAssigned : ARRAY [1..3] OF BOOL; // Дополнительный слот уже выдан типу
END_VAR
FOR uiType := UINT#1 TO UINT#3 DO
	auiMachineShare[uiType] := UINT#0;
	auiQuota[uiType] := UINT#0;
	auiRemainder[uiType] := UINT#0;
	axExtraAssigned[uiType] := FALSE;
END_FOR;

FOR uiMachine := UINT#1 TO UINT#3 DO
	IF (Config.auiMachineType[uiMachine] >= UINT#1)
	AND (Config.auiMachineType[uiMachine] <= Config.uiTypeCount) THEN
		auiMachineShare[Config.auiMachineType[uiMachine]] :=
			auiMachineShare[Config.auiMachineType[uiMachine]] + UINT#1;
	END_IF;
END_FOR;

uiAssigned := UINT#0;
FOR uiType := UINT#1 TO Config.uiTypeCount DO
	auiQuota[uiType] := (Status.uiActiveSlotCount * auiMachineShare[uiType]) / UINT#3;
	auiRemainder[uiType] := (Status.uiActiveSlotCount * auiMachineShare[uiType]) MOD UINT#3;
	uiAssigned := uiAssigned + auiQuota[uiType];
END_FOR;

uiRemaining := Status.uiActiveSlotCount - uiAssigned;
WHILE uiRemaining > UINT#0 DO
	uiBestType := UINT#0;
	uiBestRemainder := UINT#0;
	FOR uiType := UINT#1 TO Config.uiTypeCount DO
		IF NOT axExtraAssigned[uiType]
		AND ((uiBestType = UINT#0) OR (auiRemainder[uiType] > uiBestRemainder)) THEN
			uiBestType := uiType;
			uiBestRemainder := auiRemainder[uiType];
		END_IF;
	END_FOR;
	IF uiBestType = UINT#0 THEN
		uiBestType := UINT#1;
	END_IF;
	auiQuota[uiBestType] := auiQuota[uiBestType] + UINT#1;
	axExtraAssigned[uiBestType] := TRUE;
	uiRemaining := uiRemaining - UINT#1;
END_WHILE;

uiSlot := UINT#1;
FOR uiType := UINT#1 TO Config.uiTypeCount DO
	uiAssigned := UINT#0;
	WHILE (uiAssigned < auiQuota[uiType])
	AND (uiSlot <= Status.uiActiveSlotCount) DO
		Config.auiSlotType[uiSlot] := uiType;
		uiAssigned := uiAssigned + UINT#1;
		uiSlot := uiSlot + UINT#1;
	END_WHILE;
END_FOR;

FOR uiSlot := Status.uiActiveSlotCount + UINT#1 TO SINT_TO_UINT(GVL_CELL_SETTINGS.NumberDetail) DO
	Config.auiSlotType[uiSlot] := UINT#0;
END_FOR;
END_METHOD

METHOD PRIVATE RaiseWarning
VAR_INPUT
	uiCode : UINT; // Код отклонённой команды конфигурации
END_VAR
Status.stWarning.uiCode := uiCode;
Status.stWarning.udiSequence := Status.stWarning.udiSequence + UDINT#1;
IF Status.stWarning.udiSequence = UDINT#0 THEN
	Status.stWarning.udiSequence := UDINT#1;
END_IF;
END_METHOD

END_FUNCTION_BLOCK

// Device/Application/FB/FB_CELL_SAFETY
FUNCTION_BLOCK FB_CELL_SAFETY
VAR_INPUT
	axDoorLockClosedInput : ARRAY [1..4] OF BOOL;
	axDoorUnlockButtonInput : ARRAY [1..4] OF BOOL;
	axMagazineMechanismBusy : ARRAY [1..2] OF BOOL; // Только новый механизм, включая фактическое движение оси
	axEmergencyStopButtonStationInput : ARRAY [1..4] OF BOOL;
	axEmergencyStopCabinetInput : ARRAY [1..2] OF BOOL;
	xEmergencyStopMpgInput : BOOL;
	xPhaseRelayOkInput    : BOOL;
	xPressureRelayOkInput : BOOL;
	xSafetyRelayOkInput   : BOOL;
	xCellStartButtonInput : BOOL;
	xCellStopButtonInput  : BOOL;
	xCellResetButtonInput : BOOL;
	xMpgAxisXInput : BOOL;
	xMpgAxisYInput : BOOL;
	xMpgAxisZInput : BOOL;
	xMpgMultiplier1Input : BOOL;
	xMpgMultiplier10Input : BOOL;
	xMpgMultiplier100Input : BOOL;
	xSafetyRelayReset : BOOL; // Импульс отдельного сброса реле безопасности
	astMagazineStatus : ARRAY [1..2] OF ST_MAGAZINE_STATUS;
	FaultRequest : ST_CELL_SAFETY_FAULT_REQUEST;
END_VAR
VAR_OUTPUT
	Status : ST_CELL_SAFETY_STATUS;
	Error  : ST_CELL_SAFETY_ERRORS;
	Diag   : ST_CELL_SAFETY_DIAG;
	FaultStatus : ST_FAULT_INJECTION_STATUS;
	astButtonStationIoStatus : ARRAY [1..4] OF ST_BUTTON_STATION_IO_STATUS;
	stFrontControlCabinetIoStatus : ST_CONTROL_CABINET_IO_STATUS;
	stRearControlCabinetIoStatus : ST_CONTROL_CABINET_IO_STATUS;
	stMpgIoStatus : ST_MPG_IO_STATUS;
	astEnclosureDoorStatus : ARRAY [1..4] OF ST_ENCLOSURE_DOOR_STATUS;
	axDoorUnlockOutput : ARRAY [1..4] OF BOOL;
	axDoorButtonLampOutput : ARRAY [1..4] OF BOOL;
	xSafetyRelayResetOutput : BOOL;
	xCellEnablePulse : BOOL;
	xCellDisablePulse : BOOL;
	xCellResetPulse : BOOL;
END_VAR
VAR
	fbFaultInjector : FB_CELL_SAFETY_FAULT_INJECTOR;
	axEmergencyStopStation : ARRAY [1..4] OF BOOL;
	axEmergencyStopCabinet : ARRAY [1..2] OF BOOL;
	axDoorLocked : ARRAY [1..4] OF BOOL;
	axDoorUnlockDemand : ARRAY [1..4] OF BOOL;
	axDoorSeenUnlocked : ARRAY [1..4] OF BOOL;
	artDoorButton : ARRAY [1..4] OF R_TRIG;
	rtSafetyRelayReset : R_TRIG;
	tpSafetyRelayReset : TP;
	rtCellStart : R_TRIG;
	rtCellStop : R_TRIG;
	rtCellReset : R_TRIG;
	xEmergencyStopMpg : BOOL;
	xPhaseRelayOk : BOOL;
	xPressureRelayOk : BOOL;
	xSafetyRelayOk : BOOL;
	dwLiveFaultMask : DWORD;
	uiDoor : UINT;
	uiMagazine : UINT;
END_VAR
VAR CONSTANT
	ERR_ESTOP_STATION_1 : DWORD := DWORD#16#0000_0001;
	ERR_ESTOP_STATION_2 : DWORD := DWORD#16#0000_0002;
	ERR_ESTOP_STATION_3 : DWORD := DWORD#16#0000_0004;
	ERR_ESTOP_STATION_4 : DWORD := DWORD#16#0000_0008;
	ERR_ESTOP_CABINET_FRONT : DWORD := DWORD#16#0000_0010;
	ERR_ESTOP_CABINET_REAR  : DWORD := DWORD#16#0000_0020;
	ERR_ESTOP_MPG      : DWORD := DWORD#16#0000_0040;
	ERR_PHASE_RELAY    : DWORD := DWORD#16#0000_0080;
	ERR_PRESSURE_RELAY : DWORD := DWORD#16#0000_0100;
	ERR_SAFETY_RELAY   : DWORD := DWORD#16#0000_0200;
	ERR_DOOR_1_UNLOCKED : DWORD := DWORD#16#0000_0400;
	ERR_DOOR_2_UNLOCKED : DWORD := DWORD#16#0000_0800;
	ERR_DOOR_3_UNLOCKED : DWORD := DWORD#16#0000_1000;
	ERR_DOOR_4_UNLOCKED : DWORD := DWORD#16#0000_2000;
	WRN_SAFETY_RESET_REJECTED : UINT := UINT#1;
	WRN_DOOR_1_UNLOCK_REJECTED : UINT := UINT#2;
END_VAR

fbFaultInjector(Request := FaultRequest);
FaultStatus := fbFaultInjector.Status;

FOR uiDoor := UINT#1 TO UINT#4 DO
	axEmergencyStopStation[uiDoor] := axEmergencyStopButtonStationInput[uiDoor]
		OR fbFaultInjector.axEmergencyStopStation[uiDoor];
	axDoorLocked[uiDoor] := axDoorLockClosedInput[uiDoor]
		AND NOT fbFaultInjector.axDoorUnlocked[uiDoor];
	artDoorButton[uiDoor](CLK := axDoorUnlockButtonInput[uiDoor]);

	IF uiDoor <= UINT#2 THEN
		uiMagazine := UINT#1;
	ELSE
		uiMagazine := UINT#2;
	END_IF;
	astEnclosureDoorStatus[uiDoor].xUnlockAllowed := NOT astMagazineStatus[uiMagazine].xEnabled AND NOT axMagazineMechanismBusy[uiMagazine];
	axDoorButtonLampOutput[uiDoor] := astEnclosureDoorStatus[uiDoor].xUnlockAllowed;

	IF artDoorButton[uiDoor].Q THEN
		IF astEnclosureDoorStatus[uiDoor].xUnlockAllowed THEN
			axDoorUnlockDemand[uiDoor] := TRUE;
			axDoorSeenUnlocked[uiDoor] := FALSE;
		ELSE
			RaiseWarning(uiCode := WRN_DOOR_1_UNLOCK_REJECTED + uiDoor - UINT#1);
		END_IF;
	END_IF;

	// Команда держится до фактического цикла «замок открылся -> снова закрылся».
	// Если магазин включили поверх открытого доступа, выход снимается немедленно.
	IF NOT astEnclosureDoorStatus[uiDoor].xUnlockAllowed THEN
		axDoorUnlockDemand[uiDoor] := FALSE;
		axDoorSeenUnlocked[uiDoor] := FALSE;
	ELSIF axDoorUnlockDemand[uiDoor] THEN
		IF NOT axDoorLocked[uiDoor] THEN
			axDoorSeenUnlocked[uiDoor] := TRUE;
		ELSIF axDoorSeenUnlocked[uiDoor] THEN
			axDoorUnlockDemand[uiDoor] := FALSE;
			axDoorSeenUnlocked[uiDoor] := FALSE;
		END_IF;
	END_IF;

	axDoorUnlockOutput[uiDoor] := axDoorUnlockDemand[uiDoor];
	astEnclosureDoorStatus[uiDoor].xLocked := axDoorLocked[uiDoor];
	astEnclosureDoorStatus[uiDoor].xUnlockOutput := axDoorUnlockOutput[uiDoor];
	astButtonStationIoStatus[uiDoor].xEmergencyStopPressed := axEmergencyStopStation[uiDoor];
	astButtonStationIoStatus[uiDoor].xButtonPressed := axDoorUnlockButtonInput[uiDoor];
	astButtonStationIoStatus[uiDoor].xButtonLightOn := axDoorButtonLampOutput[uiDoor];
	Status.axEmergencyStopReleased[uiDoor] := NOT axEmergencyStopStation[uiDoor];
	Status.axDoorReady[uiDoor] := astEnclosureDoorStatus[uiDoor].xUnlockAllowed OR axDoorLocked[uiDoor];
	Status.axButtonStationPressed[uiDoor] := astButtonStationIoStatus[uiDoor].xButtonPressed;
	Status.axButtonStationLightOn[uiDoor] := astButtonStationIoStatus[uiDoor].xButtonLightOn;
END_FOR;

FOR uiDoor := UINT#1 TO UINT#2 DO
	axEmergencyStopCabinet[uiDoor] := axEmergencyStopCabinetInput[uiDoor]
		OR fbFaultInjector.axEmergencyStopCabinet[uiDoor];
	Status.axEmergencyStopReleased[uiDoor + UINT#4] := NOT axEmergencyStopCabinet[uiDoor];
END_FOR;
xEmergencyStopMpg := xEmergencyStopMpgInput OR fbFaultInjector.xEmergencyStopMpg;
Status.axEmergencyStopReleased[7] := NOT xEmergencyStopMpg;

xPhaseRelayOk := xPhaseRelayOkInput AND NOT fbFaultInjector.xPhaseRelayFault;
xPressureRelayOk := xPressureRelayOkInput AND NOT fbFaultInjector.xPressureRelayFault;
xSafetyRelayOk := xSafetyRelayOkInput AND NOT fbFaultInjector.xSafetyRelayFault;

rtSafetyRelayReset(CLK := xSafetyRelayReset);
Status.xSafetyRelayResetAllowed := NOT xSafetyRelayOk AND NOT tpSafetyRelayReset.Q;
IF rtSafetyRelayReset.Q AND NOT Status.xSafetyRelayResetAllowed THEN
	RaiseWarning(uiCode := WRN_SAFETY_RESET_REJECTED);
END_IF;
tpSafetyRelayReset(
	IN := rtSafetyRelayReset.Q AND Status.xSafetyRelayResetAllowed,
	PT := T#1S
);
// Разрешение проверяется на фронте команды; после запуска выдаём полный импульс 1 с.
xSafetyRelayResetOutput := tpSafetyRelayReset.Q;
Status.xSafetyRelayResetActive := xSafetyRelayResetOutput;

rtCellStart(CLK := xCellStartButtonInput);
rtCellStop(CLK := xCellStopButtonInput);
rtCellReset(CLK := xCellResetButtonInput);
xCellEnablePulse := rtCellStart.Q;
xCellDisablePulse := rtCellStop.Q;
xCellResetPulse := rtCellReset.Q;

stFrontControlCabinetIoStatus.xEmergencyStopPressed := axEmergencyStopCabinet[1];
stFrontControlCabinetIoStatus.xStartPressed := xCellStartButtonInput;
stFrontControlCabinetIoStatus.xStopPressed := xCellStopButtonInput;
stFrontControlCabinetIoStatus.xResetPressed := xCellResetButtonInput;
stRearControlCabinetIoStatus.xEmergencyStopPressed := axEmergencyStopCabinet[2];
stRearControlCabinetIoStatus.xStartPressed := FALSE;
stRearControlCabinetIoStatus.xStopPressed := FALSE;
stRearControlCabinetIoStatus.xResetPressed := FALSE;
stMpgIoStatus.xEmergencyStopPressed := xEmergencyStopMpg;
stMpgIoStatus.xAxisX := xMpgAxisXInput;
stMpgIoStatus.xAxisY := xMpgAxisYInput;
stMpgIoStatus.xAxisZ := xMpgAxisZInput;
stMpgIoStatus.xMultiplier1 := xMpgMultiplier1Input;
stMpgIoStatus.xMultiplier10 := xMpgMultiplier10Input;
stMpgIoStatus.xMultiplier100 := xMpgMultiplier100Input;

dwLiveFaultMask := DWORD#0;
IF axEmergencyStopStation[1] THEN dwLiveFaultMask := dwLiveFaultMask OR ERR_ESTOP_STATION_1; END_IF;
IF axEmergencyStopStation[2] THEN dwLiveFaultMask := dwLiveFaultMask OR ERR_ESTOP_STATION_2; END_IF;
IF axEmergencyStopStation[3] THEN dwLiveFaultMask := dwLiveFaultMask OR ERR_ESTOP_STATION_3; END_IF;
IF axEmergencyStopStation[4] THEN dwLiveFaultMask := dwLiveFaultMask OR ERR_ESTOP_STATION_4; END_IF;
IF axEmergencyStopCabinet[1] THEN dwLiveFaultMask := dwLiveFaultMask OR ERR_ESTOP_CABINET_FRONT; END_IF;
IF axEmergencyStopCabinet[2] THEN dwLiveFaultMask := dwLiveFaultMask OR ERR_ESTOP_CABINET_REAR; END_IF;
IF xEmergencyStopMpg THEN dwLiveFaultMask := dwLiveFaultMask OR ERR_ESTOP_MPG; END_IF;
IF NOT xPhaseRelayOk THEN dwLiveFaultMask := dwLiveFaultMask OR ERR_PHASE_RELAY; END_IF;
IF NOT xPressureRelayOk THEN dwLiveFaultMask := dwLiveFaultMask OR ERR_PRESSURE_RELAY; END_IF;
IF NOT xSafetyRelayOk THEN dwLiveFaultMask := dwLiveFaultMask OR ERR_SAFETY_RELAY; END_IF;
IF (astMagazineStatus[1].xEnabled OR axMagazineMechanismBusy[1]) AND NOT axDoorLocked[1] THEN dwLiveFaultMask := dwLiveFaultMask OR ERR_DOOR_1_UNLOCKED; END_IF;
IF (astMagazineStatus[1].xEnabled OR axMagazineMechanismBusy[1]) AND NOT axDoorLocked[2] THEN dwLiveFaultMask := dwLiveFaultMask OR ERR_DOOR_2_UNLOCKED; END_IF;
IF (astMagazineStatus[2].xEnabled OR axMagazineMechanismBusy[2]) AND NOT axDoorLocked[3] THEN dwLiveFaultMask := dwLiveFaultMask OR ERR_DOOR_3_UNLOCKED; END_IF;
IF (astMagazineStatus[2].xEnabled OR axMagazineMechanismBusy[2]) AND NOT axDoorLocked[4] THEN dwLiveFaultMask := dwLiveFaultMask OR ERR_DOOR_4_UNLOCKED; END_IF;

Error.dwErrorActive := dwLiveFaultMask;
Error.dwAlarmActive := dwLiveFaultMask;
IF dwLiveFaultMask <> DWORD#0 THEN
	Error.dwErrorLast := dwLiveFaultMask;
END_IF;
Status.xPhaseRelayOk := xPhaseRelayOk;
Status.xPressureRelayOk := xPressureRelayOk;
Status.xSafetyRelayOk := xSafetyRelayOk;
Status.xGlobalError := dwLiveFaultMask <> DWORD#0;
Status.xReady := NOT Status.xGlobalError;

METHOD PRIVATE RaiseWarning
VAR_INPUT
	uiCode : UINT;
END_VAR
Diag.stWarning.uiCode := uiCode;
Diag.stWarning.udiSequence := Diag.stWarning.udiSequence + UDINT#1;
IF Diag.stWarning.udiSequence = UDINT#0 THEN
	Diag.stWarning.udiSequence := UDINT#1;
END_IF;
END_METHOD

END_FUNCTION_BLOCK

// Device/Application/FB/FB_FAULT_INJECTOR/FB_CELL_SAFETY_FAULT_INJECTOR
FUNCTION_BLOCK FB_CELL_SAFETY_FAULT_INJECTOR
VAR_INPUT
	Request : ST_CELL_SAFETY_FAULT_REQUEST;
END_VAR
VAR_OUTPUT
	axEmergencyStopStation : ARRAY [1..4] OF BOOL;
	axEmergencyStopCabinet : ARRAY [1..2] OF BOOL;
	xEmergencyStopMpg   : BOOL;
	xPhaseRelayFault    : BOOL;
	xPressureRelayFault : BOOL;
	xSafetyRelayFault   : BOOL;
	axDoorUnlocked      : ARRAY [1..4] OF BOOL;
	Status              : ST_FAULT_INJECTION_STATUS;
END_VAR
VAR
	uiIndex : UINT;
END_VAR

Status.xAllowed := Request.xEnabled;
Status.xBusy := FALSE;
Status.xRejected := FALSE;
Status.xResetAllowed := FALSE;

FOR uiIndex := UINT#1 TO UINT#4 DO
	axEmergencyStopStation[uiIndex] := Request.xEnabled AND Request.axEmergencyStopStation[uiIndex];
	axDoorUnlocked[uiIndex] := Request.xEnabled AND Request.axDoorUnlocked[uiIndex];
END_FOR;
FOR uiIndex := UINT#1 TO UINT#2 DO
	axEmergencyStopCabinet[uiIndex] := Request.xEnabled AND Request.axEmergencyStopCabinet[uiIndex];
END_FOR;
xEmergencyStopMpg := Request.xEnabled AND Request.xEmergencyStopMpg;
xPhaseRelayFault := Request.xEnabled AND Request.xPhaseRelayFault;
xPressureRelayFault := Request.xEnabled AND Request.xPressureRelayFault;
xSafetyRelayFault := Request.xEnabled AND Request.xSafetyRelayFault;

Status.xActive := xEmergencyStopMpg
	OR xPhaseRelayFault
	OR xPressureRelayFault
	OR xSafetyRelayFault;
FOR uiIndex := UINT#1 TO UINT#4 DO
	Status.xActive := Status.xActive
		OR axEmergencyStopStation[uiIndex]
		OR axDoorUnlocked[uiIndex];
END_FOR;
FOR uiIndex := UINT#1 TO UINT#2 DO
	Status.xActive := Status.xActive OR axEmergencyStopCabinet[uiIndex];
END_FOR;

END_FUNCTION_BLOCK

// Device/Application/FB/FB_CELL_MANAGER/FB_CELL_MANAGER
FUNCTION_BLOCK FB_CELL_MANAGER
VAR_INPUT
	xIoManual : BOOL; // Прямой ручной слой отменяет задание, не сбрасывая аварии
	axMagazineAutoSwapPending : ARRAY [1..GVL_CELL_SETTINGS.MagazineCount] OF BOOL; // Палета ждёт окна обмена
	axMagazineExchangeInProgress : ARRAY [1..GVL_CELL_SETTINGS.MagazineCount] OF BOOL; // Во время смены палет запрещены операции только с этим магазином
	xMagazineExchangeActive : BOOL; // Есть активный обмен палет; подавляет временные предупреждения о запасах
	xStart            : BOOL; // Импульс запуска цикла или отмены остановки
	xStop             : BOOL; // Импульс контролируемой остановки
	xTestAbort        : BOOL; // Немедленная отмена только тестового прогона
	xResetRequest     : BOOL; // Необработанный запрос сброса от HMI
	xReset            : BOOL; // Общий сброс владельцев ошибок
	xOperatorChoice   : BOOL; // Импульс ответа активному предпусковому опросу
	xOperatorCancel   : BOOL; // Импульс отмены предпускового опроса
	uiOperatorChoice  : UINT; // Выбранное содержимое, тип продукции или станок
	xManual           : BOOL; // Ручной режим ячейки
	xIoDoRejected : BOOL;
    xIoEmergencyResetRejected : BOOL;
    xIoEmergencyStopActive : BOOL;
	xIoOverrideRejected : BOOL; // Отклонённая транзакция диагностики, эффект WARNING
	xSettingsRejected : BOOL; // Rejected or expired setting transaction
	uiModeRejectReason : UINT; // Одноцикловый отказ транзакции режима: 2 цикл, 3 Safety
	xGlobalError      : BOOL; // Глобальная ошибка ячейки
	xSafetyReady      : BOOL; // Все дискретные условия безопасности выполнены
	xDrivesReady      : BOOL; // Приводы готовы
	xMotionBusy       : BOOL; // Оси ещё движутся
	xRobotInterfaceReady : BOOL; // Выбранный интерфейс робота готов к работе
	lrRobotActualX    : LREAL; // Фактическая координата робота X
	lrRobotActualY    : LREAL; // Фактическая координата робота Y
	lrRobotActualZ    : LREAL; // Фактическая координата робота Z
	stSafetyHomePoint : ST_POINT; // Настроенная безопасная точка повторного запуска
	lrSafetyHomeToleranceX : LREAL; // Допуск HOME_SAFETY по X
	lrSafetyHomeToleranceY : LREAL; // Допуск HOME_SAFETY по Y
	lrSafetyHomeToleranceZ : LREAL; // Допуск HOME_SAFETY по Z
	lrStoppedPoseTolerance : LREAL; // Допуск контроля позы после штатной остановки
	Config            : ST_MULTI_TYPE_CONFIG; // Активная конфигурация типов
	xConfigurationValid : BOOL; // Конфигурация типов прошла проверку
	xPointsConfigured : BOOL; // HOME_SAFETY и точки включённого оборудования настроены
	stRobotStatus     : ST_ROBOT_STATUS; // Состояние робота
	astMagazineStatus : ARRAY [1..GVL_CELL_SETTINGS.MagazineCount] OF ST_MAGAZINE_STATUS;
	astMachineStatus  : ARRAY [1..3] OF ST_MACHINE_PUBLIC; // Состояния станков
	astMachineDiag    : ARRAY [1..3] OF ST_MACHINE_DIAG; // Автоматы станков
	FaultRequest      : ST_CELL_FAULT_REQUEST; // Диагностическая инъекция
END_VAR
VAR_OUTPUT
	Command            : ST_CELL_COMMAND; // Команды существующим блокам ячейки
	Status             : ST_CELL_STATUS; // Общий контракт состояния ячейки
	Diag               : ST_CELL_DIAG; // Общий контракт диагностики ячейки
	Error              : ST_CELL_ERRORS; // Общий контракт ошибок ячейки
	CycleStatus        : ST_CELL_CYCLE_STATUS; // Расширенная диагностика универсального цикла
	FaultStatus        : ST_FAULT_INJECTION_STATUS; // Инъекция логической ошибки ячейки
END_VAR
VAR
	axGeometryUnloadBlocked : ARRAY [1..3] OF BOOL; // Вызванная деталь ждёт свободного ГК или своей очереди FIFO
	atonGeometryWait : ARRAY [1..3] OF TON;
	audiGeometryWaitCallId : ARRAY [1..3] OF UDINT;
	axGeometryWaitWarned : ARRAY [1..3] OF BOOL;
	xGeometryHeld : BOOL;
	xGeometryDetailCounted : BOOL;
	uiGeometryMachine : UINT;
	uiGeometryStation : UINT;
	uiGeometryParkStation : UINT;
	uiGeometryStep : UINT;
	uiGeometryBypassReason : UINT;
	uiGeometryIndex : UINT;
	udiGeometryMagazineCounter : UDINT;
	eGeometryReturnState : E_CELL_MANAGER_STATE;
	eGeometrySafePoint : E_POINT_NAME;
	eGeometryChangePoint : E_POINT_NAME;
	eGeometryPlacePoint : E_POINT_NAME;
	xActiveMagazineAutoSwapPending : BOOL; // Удержать владельца и цикл до обмена его палеты
	eState               : E_CELL_MANAGER_STATE := E_CELL_MANAGER_STATE.IDLE; // Состояние универсального автомата
	eMagazineOperation   : E_MAGAZINE_OPERATION; // Выполняемая операция магазина
	eMachineOperation    : E_MACHINE_OPERATION; // Зафиксированная операция станка
	xRunning             : BOOL; // Защёлка автоматического цикла
	xStopRequested       : BOOL; // Остановка после безопасного шага
	xReadyToStart        : BOOL; // Условия запуска выполнены
	xRobotReady          : BOOL; // Робот готов принять маршрут
	xMagazineReady       : BOOL; // Магазин готов к операции
	xActiveMagazineExchangeInProgress : BOOL; // Выбранный магазин сейчас меняет палеты
	stMagazineStatus     : ST_MAGAZINE_STATUS; // Снимок выбранного магазина для существующего автомата
	uiActiveMagazine     : UINT; // Защёлкнутый магазин текущего цикла
	xMagazine1Available  : BOOL;
	xMagazine2Available  : BOOL;
	xMagazineSelectionAllowed : BOOL; // Новое владение допускается только между операциями
	xMagazine1CanContinue : BOOL; // Первый магазин позволяет следующий технологический шаг
	xMagazine2CanContinue : BOOL; // Второй магазин позволяет следующий технологический шаг
	xMagazine1CanSupplyBlank : BOOL; // М1 позволяет штатный план TAKE перед отдельной выгрузкой
	xMagazine2CanSupplyBlank : BOOL; // М2 позволяет штатный план TAKE перед отдельной выгрузкой
	xMagazine1CanExchangeDetail : BOOL; // Заготовка М1 освобождает слот для детали робота
	xMagazine2CanExchangeDetail : BOOL;
	xActiveMagazineCanExchangeDetail : BOOL;
	xHeldBlankLoadAvailable : BOOL; // При двух грузах можно сначала загрузить пустой станок
	xMagazineMachineWorkPending : BOOL; // Из станка ещё потребуется выгрузка
	uiMagazineType       : UINT; // Тип станка при проверке содержимого обоих магазинов
	uiPreferredMagazine  : UINT; // Первый подходящий магазин в порядке 1, 2
	xReselectMagazine    : BOOL; // Требуется передать владение подходящему магазину
	xAlternateMagazineAvailable : BOOL; // Второй магазин готов принять непрерывный автоматический цикл
	xUseAlternateMagazineForDetail : BOOL; // У текущего магазина нет слота детали, у второго есть
	xAnyMagazineDetailSlotAvailable : BOOL; // Есть доступный слот детали хотя бы в одном магазине
	xNoDetailDestinationCondition : BOOL; // Робот держит готовую деталь без доступного слота
	xNoBlankStockCondition : BOOL; // Нет заготовок и текущей работы для автоматического цикла
	xDetailDestinationWarningActive : BOOL; // Предупреждение об отсутствии места уже выдано
	xBlankStockWarningActive : BOOL; // Предупреждение об отсутствии заготовок уже выдано
	xMachineWorkPending : BOOL; // Станок занят/обрабатывает, запускается или содержит изделие
	xAnyMachineBusy      : BOOL; // Хотя бы один станок обслуживается
	xMachineServiceStarted : BOOL; // Выбранный станок вошёл в рецепт
	xReselectAfterRobotRelease : BOOL; // После снятия команды требуется повторный выбор
	xChangePrepared      : BOOL; // Для CHANGE зафиксированы совместимый станок и два корректных слота
	xFaultAllowed        : BOOL; // Инъекция разрешена в полностью остановленной ячейке
	xResetAllowed        : BOOL; // Локальная ошибка может быть сброшена
	xPayloadRouteWarningActive : BOOL; // Предупреждение о несовпадении типа груза и назначения уже выдано
	xPrestartGripper1Occupied : BOOL; // Снимок занятости первого захвата на момент запуска опроса
	xPrestartGripper2Occupied : BOOL; // Снимок занятости второго захвата на момент запуска опроса
	xSafetyHomeRequired : BOOL; // Защёлка обязательного возврата в HOME_SAFETY
	xRobotAtSafetyHome  : BOOL; // Робот находится в допустимом диапазоне HOME_SAFETY
	xStoppedPoseValid   : BOOL; // После штатной остановки сохранена доверенная поза
	xWasRunning         : BOOL; // Состояние цикла на предыдущем вызове
	xStartCheckCellIdle           : BOOL; // Отдельные условия запуска для HMI
	xStartCheckAutomaticMode      : BOOL;
	xStartCheckNoBlockingError    : BOOL;
	xStartCheckRobotInterfaceReady: BOOL;
	xStartCheckConfigurationValid : BOOL;
	xStartCheckPointsConfigured   : BOOL;
	xStartCheckDrivesReady        : BOOL;
	xStartCheckRobotReady         : BOOL;
	xStartCheckMagazineReady      : BOOL;
	xStartCheckTaskAvailable      : BOOL;
	xStartCheckSafetyHome         : BOOL;
	xStartCheckSafety             : BOOL;
	xOperatorPromptState          : BOOL; // Текущий шаг ожидает ответ HMI
	xOperatorChoiceAllowed        : BOOL;
	xOperatorCancelAllowed        : BOOL;
	uiOperatorPrompt              : UINT;
	uiOperatorTypeMask            : UINT;
	uiOperatorMachineMask         : UINT;
	uiStartConditionsMet         : UINT;
	lrStoppedPoseX      : LREAL; // Доверенная координата X штатной остановки
	lrStoppedPoseY      : LREAL; // Доверенная координата Y штатной остановки
	lrStoppedPoseZ      : LREAL; // Доверенная координата Z штатной остановки
	uiReadyMachines      : UINT; // Число доступных маршрутных целей
	uiMachine            : UINT; // Индекс станка
	uiMagazineIndex      : UINT; // Индекс магазина при поиске свободного слота
	uiCandidateMachine   : UINT; // Результат выбора
	uiSelectedMachine    : UINT; // Зафиксированный станок
	uiSelectedType       : UINT; // Тип маршрута
	uiBlankPayloadType   : UINT; // Тип заготовки в первом захвате
	uiDetailPayloadType  : UINT; // Тип готовой детали во втором захвате
	axMachineStartPending: ARRAY [1..3] OF BOOL; // Станок обслужен, но xProcessing ещё не подтверждён
	iTakeSlot            : SINT; // Зарезервированный слот заготовки
	iPutSlot             : SINT; // Зарезервированный слот укладки
	iTakeOriginSlot      : SINT; // Исходный слот заготовки для приоритетного возврата
	rtStart              : R_TRIG; // Фронт запуска
	rtStop               : R_TRIG; // Фронт остановки
	rtReset              : R_TRIG; // Фронт сброса
	rtOperatorChoice     : R_TRIG; // Один ответ не переносится на следующий шаг опроса
	rtOperatorCancel     : R_TRIG; // Фронт отмены предпускового опроса
	fbFaultInjector      : FB_CELL_FAULT_INJECTOR; // Проверка противоречивого груза
END_VAR
VAR CONSTANT
	FIRST_MACHINE     : UINT := UINT#1;
	LAST_MACHINE      : UINT := UINT#3;
	MACHINE_SWITCH_DEADBAND : TIME := T#1S; // Минимальный выигрыш времени для смены ожидаемой цели
	START_PENDING_ESTIMATE  : TIME := T#1S; // Оценка перехода от освобождения робота до xProcessing
	ERR_BOTH_GRIPPERS : DWORD := DWORD#16#0000_0001;
	ERR_ROBOT         : DWORD := DWORD#16#0000_0002;
	ERR_MAGAZINE      : DWORD := DWORD#16#0000_0004;
	ERR_MACHINE       : DWORD := DWORD#16#0000_0008;
	ERR_GLOBAL_STOP   : DWORD := DWORD#16#0000_0010;
	WRN_START_NOT_READY       : UINT := UINT#4;
	WRN_STOP_NOT_RUNNING      : UINT := UINT#5;
	WRN_SIM_ERROR_NOT_ALLOWED : UINT := UINT#8;
	WRN_PAYLOAD_ROUTE_MISMATCH : UINT := UINT#9;
	WRN_SAFETY_HOME_REQUIRED   : UINT := UINT#10;
	WRN_MANUAL_MODE_REJECTED   : UINT := UINT#11;
	WRN_CELL_SETTING_REJECTED : UINT := UINT#28;
	WRN_AUTOMATIC_MODE_REJECTED : UINT := UINT#27; // WARNING: общая авария удерживает ручной режим
	WRN_GRIPPER1_CONTENT       : UINT := UINT#15;
	WRN_GRIPPER2_CONTENT       : UINT := UINT#16;
	WRN_PAYLOAD_TYPE_CHOICE    : UINT := UINT#17;
	WRN_DETAIL_SLOT_REQUIRED   : UINT := UINT#18;
	WRN_START_MACHINE_REQUIRED : UINT := UINT#19;
	WRN_START_MACHINE_CHOICE   : UINT := UINT#20;
	WRN_OPERATOR_REPLY_REJECTED: UINT := UINT#21;
	WRN_OPERATOR_CANCEL_REJECTED: UINT := UINT#22;
	WRN_NO_DETAIL_DESTINATION  : UINT := UINT#29;
	WRN_NO_BLANK_STOCK         : UINT := UINT#30;
	WRN_GEOMETRY_WAIT_TIMEOUT  : UINT := UINT#52;
	WRN_IO_OVERRIDE_REJECTED   : UINT := UINT#31;
    WRN_IO_DO_REJECTED : UINT := UINT#32;
    WRN_IO_EMERGENCY_RESET_REJECTED : UINT := UINT#33;
END_VAR

IF xIoDoRejected THEN
    Diag.stWarning.uiCode := WRN_IO_DO_REJECTED; // WARNING: вход/команда прямого ручного I/O не применены
    Diag.stWarning.udiSequence := Diag.stWarning.udiSequence + UDINT#1;
    IF Diag.stWarning.udiSequence = UDINT#0 THEN Diag.stWarning.udiSequence := UDINT#1; END_IF;
END_IF;
IF xIoEmergencyResetRejected THEN
    Diag.stWarning.uiCode := WRN_IO_EMERGENCY_RESET_REJECTED; // WARNING: останов остаётся
    Diag.stWarning.udiSequence := Diag.stWarning.udiSequence + UDINT#1;
    IF Diag.stWarning.udiSequence = UDINT#0 THEN Diag.stWarning.udiSequence := UDINT#1; END_IF;
END_IF;
IF xIoOverrideRejected THEN
    Diag.stWarning.uiCode := WRN_IO_OVERRIDE_REJECTED; // WARNING: входы не изменены
    Diag.stWarning.udiSequence := Diag.stWarning.udiSequence + UDINT#1;
    IF Diag.stWarning.udiSequence = UDINT#0 THEN Diag.stWarning.udiSequence := UDINT#1; END_IF;
END_IF;
IF xSettingsRejected THEN
	Diag.stWarning.uiCode := WRN_CELL_SETTING_REJECTED; // WARNING: settings unchanged
	Diag.stWarning.udiSequence := Diag.stWarning.udiSequence + UDINT#1;
	IF Diag.stWarning.udiSequence = UDINT#0 THEN Diag.stWarning.udiSequence := UDINT#1; END_IF;
END_IF;


rtStart(CLK := xStart);
rtStop(CLK := xStop);
rtReset(CLK := xResetRequest);
rtOperatorChoice(CLK := xOperatorChoice);
rtOperatorCancel(CLK := xOperatorCancel);

// До выбора магазина/станка исключаем выгрузку вызванной детали без свободного ГК.
UpdateGeometryWait();

// Выбор выполняется только между операциями. Внутренний автомат по-прежнему
// работает с одним снимком, поэтому уже отлажанный маршрут не размазывается
// по двум владельцам и не переключается посреди TAKE/CHANGE.
xMagazine1Available := astMagazineStatus[1].xEnabled
	AND astMagazineStatus[1].xReady
	AND NOT axMagazineExchangeInProgress[1]
	AND NOT astMagazineStatus[1].xBusy
	AND NOT astMagazineStatus[1].xError
	AND NOT astMagazineStatus[1].xDisablePending
	AND NOT astMagazineStatus[1].xFinished;
xMagazine2Available := astMagazineStatus[2].xEnabled
	AND astMagazineStatus[2].xReady
	AND NOT axMagazineExchangeInProgress[2]
	AND NOT astMagazineStatus[2].xBusy
	AND NOT astMagazineStatus[2].xError
	AND NOT astMagazineStatus[2].xDisablePending
	AND NOT astMagazineStatus[2].xFinished;

// Полная палета тоже принимает деталь: сначала берём заготовку свободным
// захватом 1, затем кладём деталь в освободившийся универсальный слот.
// Заготовке нужен совместимый маршрут; станок может ещё обрабатывать изделие.
xMagazine1CanExchangeDetail := FALSE;
xMagazine2CanExchangeDetail := FALSE;
xHeldBlankLoadAvailable := FALSE;
FOR uiMachine := FIRST_MACHINE TO LAST_MACHINE DO
	IF IsMachineEligible(uiMachine := uiMachine) THEN
		uiMagazineType := Config.auiMachineType[uiMachine];
		IF stRobotStatus.xBlankAvailable AND stRobotStatus.xDetailAvailable
		AND (uiMagazineType = uiBlankPayloadType)
		AND astMachineStatus[uiMachine].xCanAcceptService
		AND (astMachineStatus[uiMachine].ePartState = E_PART_STATE.EMPTY) THEN
			xHeldBlankLoadAvailable := TRUE;
		END_IF;
		IF stRobotStatus.xDetailAvailable
		AND NOT stRobotStatus.xBlankAvailable
		AND stRobotStatus.xGripper1Open
		AND (uiDetailPayloadType >= UINT#1)
		AND (uiDetailPayloadType <= Config.uiTypeCount)
		AND (uiMagazineType >= UINT#1) AND (uiMagazineType <= UINT#3)
		AND (astMachineStatus[uiMachine].xProcessing
			OR axMachineStartPending[uiMachine]
			OR (astMachineStatus[uiMachine].xCanAcceptService
				AND ((astMachineStatus[uiMachine].ePartState = E_PART_STATE.EMPTY)
					OR astMachineStatus[uiMachine].xServiceRequired))) THEN
			IF astMagazineStatus[1].stTypeStatus.aiBlankSlot[uiMagazineType] > SINT#0 THEN
				xMagazine1CanExchangeDetail := xMagazine1Available;
			END_IF;
			IF astMagazineStatus[2].stTypeStatus.aiBlankSlot[uiMagazineType] > SINT#0 THEN
				xMagazine2CanExchangeDetail := xMagazine2Available;
			END_IF;
		END_IF;
	END_IF;
END_FOR;

// После полной выработки или операторского запроса отключения активного магазина
// автомат не требует нового Start. Переключение выполняется только когда робот
// и старый магазин уже освобождены.
xAlternateMagazineAvailable := FALSE;
IF uiActiveMagazine = UINT#1 THEN
	xAlternateMagazineAvailable := xMagazine2Available;
ELSIF uiActiveMagazine = UINT#2 THEN
	xAlternateMagazineAvailable := xMagazine1Available;
END_IF;

// Если деталь уже у робота, сначала переключаем владение на второй магазин,
// если там есть совместимый свободный слот. Это происходит только на границе
// операций и не прерывает уже выданную команду.
xUseAlternateMagazineForDetail := FALSE;
IF xRunning
AND stRobotStatus.xDetailAvailable
AND ((eState = E_CELL_MANAGER_STATE.PLAN_TARGET)
	OR (eState = E_CELL_MANAGER_STATE.WAIT_TARGET)
	OR (eState = E_CELL_MANAGER_STATE.SELECT_FALLBACK)
	OR (eState = E_CELL_MANAGER_STATE.WAIT_MAGAZINE))
AND (uiDetailPayloadType >= UINT#1)
AND (uiDetailPayloadType <= Config.uiTypeCount) THEN
	IF uiActiveMagazine = UINT#1 THEN
		IF (astMagazineStatus[1].stTypeStatus.aiFreeSlot[uiDetailPayloadType] = SINT#0)
		AND NOT xMagazine1CanExchangeDetail
		AND xMagazine2Available THEN
			IF astMagazineStatus[2].stTypeStatus.aiFreeSlot[uiDetailPayloadType] > SINT#0 THEN
				xUseAlternateMagazineForDetail := TRUE;
			END_IF;
		END_IF;
	ELSIF uiActiveMagazine = UINT#2 THEN
		IF (astMagazineStatus[2].stTypeStatus.aiFreeSlot[uiDetailPayloadType] = SINT#0)
		AND NOT xMagazine2CanExchangeDetail
		AND xMagazine1Available THEN
			IF astMagazineStatus[1].stTypeStatus.aiFreeSlot[uiDetailPayloadType] > SINT#0 THEN
				xUseAlternateMagazineForDetail := TRUE;
			END_IF;
		END_IF;
	END_IF;
END_IF;
// На каждой границе планирования проверяем ОБА магазина. Готовность механики
// сама по себе не означает наличие следующей операции: учитываем типы заготовок
// и возможность вернуть изделие из включённого исправного станка.
// Уже взятую заготовку сначала обслуживаем или возвращаем в исходный слот.
xMagazineSelectionAllowed := NOT stRobotStatus.xBusy
	AND NOT stRobotStatus.xBlankAvailable
	AND ((eState = E_CELL_MANAGER_STATE.IDLE)
		OR (eState = E_CELL_MANAGER_STATE.PLAN_TARGET)
		OR (eState = E_CELL_MANAGER_STATE.WAIT_TARGET)
		OR (eState = E_CELL_MANAGER_STATE.SELECT_FALLBACK)
		OR (eState = E_CELL_MANAGER_STATE.WAIT_MAGAZINE));
xMagazine1CanContinue := xMagazine1Available;
xMagazine2CanContinue := xMagazine2Available;
xMagazine1CanSupplyBlank := FALSE;
xMagazine2CanSupplyBlank := FALSE;
IF xRunning AND xMagazineSelectionAllowed THEN
	xMagazine1CanContinue := FALSE;
	xMagazine2CanContinue := FALSE;
	IF stRobotStatus.xDetailAvailable THEN
		IF (uiDetailPayloadType >= UINT#1)
		AND (uiDetailPayloadType <= Config.uiTypeCount)
		AND (uiDetailPayloadType <= UINT#3) THEN
			xMagazine1CanContinue := xMagazine1Available
				AND ((astMagazineStatus[1].stTypeStatus.aiFreeSlot[uiDetailPayloadType] > SINT#0)
					OR xMagazine1CanExchangeDetail);
			xMagazine2CanContinue := xMagazine2Available
				AND ((astMagazineStatus[2].stTypeStatus.aiFreeSlot[uiDetailPayloadType] > SINT#0)
					OR xMagazine2CanExchangeDetail);
		END_IF;
	ELSE
		FOR uiMachine := FIRST_MACHINE TO LAST_MACHINE DO
			IF IsMachineEligible(uiMachine := uiMachine) THEN
				uiMagazineType := Config.auiMachineType[uiMachine];
				IF (uiMagazineType >= UINT#1) AND (uiMagazineType <= UINT#3) THEN
					xMagazineMachineWorkPending := astMachineStatus[uiMachine].xProcessing
						OR axMachineStartPending[uiMachine]
						OR ((astMachineStatus[uiMachine].ePartState = E_PART_STATE.LOADED)
							AND ((astMachineStatus[uiMachine].ePartType = E_PART_TYPE.PART)
								OR (astMachineStatus[uiMachine].ePartType = E_PART_TYPE.DETAIL)));
					IF (astMagazineStatus[1].stTypeStatus.aiBlankSlot[uiMagazineType] > SINT#0)
					AND (astMachineStatus[uiMachine].xCanAcceptService OR xMagazineMachineWorkPending) THEN
						xMagazine1CanSupplyBlank := xMagazine1Available;
					END_IF;
					IF ((astMagazineStatus[1].stTypeStatus.aiBlankSlot[uiMagazineType] > SINT#0)
						AND (astMachineStatus[uiMachine].xCanAcceptService OR xMagazineMachineWorkPending))
					OR ((astMagazineStatus[1].stTypeStatus.aiFreeSlot[uiMagazineType] > SINT#0)
						AND xMagazineMachineWorkPending) THEN
						xMagazine1CanContinue := xMagazine1Available;
					END_IF;
					IF (astMagazineStatus[2].stTypeStatus.aiBlankSlot[uiMagazineType] > SINT#0)
					AND (astMachineStatus[uiMachine].xCanAcceptService OR xMagazineMachineWorkPending) THEN
						xMagazine2CanSupplyBlank := xMagazine2Available;
					END_IF;
					IF ((astMagazineStatus[2].stTypeStatus.aiBlankSlot[uiMagazineType] > SINT#0)
						AND (astMachineStatus[uiMachine].xCanAcceptService OR xMagazineMachineWorkPending))
					OR ((astMagazineStatus[2].stTypeStatus.aiFreeSlot[uiMagazineType] > SINT#0)
						AND xMagazineMachineWorkPending) THEN
						xMagazine2CanContinue := xMagazine2Available;
					END_IF;
				END_IF;
			END_IF;
		END_FOR;
	END_IF;
END_IF;
// Как и штатный PLAN_TARGET, сначала ищем TAKE, затем отдельную выгрузку.
// Пустой М1 не должен заставлять ждать обработку, если М2 позволяет загрузку.
uiPreferredMagazine := UINT#0;
IF xMagazine1CanSupplyBlank THEN
	uiPreferredMagazine := UINT#1;
ELSIF xMagazine2CanSupplyBlank THEN
	uiPreferredMagazine := UINT#2;
ELSIF xMagazine1CanContinue THEN
	uiPreferredMagazine := UINT#1;
ELSIF xMagazine2CanContinue THEN
	uiPreferredMagazine := UINT#2;
END_IF;
xReselectMagazine := xMagazineSelectionAllowed
	AND (uiPreferredMagazine > UINT#0)
	AND (uiActiveMagazine <> uiPreferredMagazine)
	AND NOT ((uiActiveMagazine = UINT#1) AND astMagazineStatus[1].xBusy)
	AND NOT ((uiActiveMagazine = UINT#2) AND astMagazineStatus[2].xBusy);

IF xRunning
AND (eState <> E_CELL_MANAGER_STATE.GEOMETRY_WAIT_FREE)
AND (eState <> E_CELL_MANAGER_STATE.GEOMETRY_DELIVER)
AND (eState <> E_CELL_MANAGER_STATE.GEOMETRY_RELEASE_COMMAND)
AND (uiActiveMagazine >= UINT#1)
AND (uiActiveMagazine <= UINT#2) THEN
	// Операторское отключение активного магазина передаёт владение второму
	// только на границе операций. Фактический груз FB_ROBOT при этом остаётся
	// источником истины и будет уложен уже в выбранный магазин. Проверяем также
	// итоговый xEnabled: FB_MAGAZINE может завершить отключение и снять
	// xDisablePending раньше, чем робот достигнет границы перепланирования.
	// xFinished в DONE ещё не означает конец цикла: до завершения RELEASE_MAGAZINE
	// не меняем владельца. Когда началась сама смена палет, адресная блокировка
	// снимает старого владельца на границе операций и разрешает выбрать второй магазин.
	IF (((astMagazineStatus[uiActiveMagazine].xFinished
			AND NOT axMagazineAutoSwapPending[uiActiveMagazine])
		OR ((astMagazineStatus[uiActiveMagazine].xDisablePending
			OR NOT astMagazineStatus[uiActiveMagazine].xEnabled)
			AND ((eState = E_CELL_MANAGER_STATE.PLAN_TARGET)
				OR (eState = E_CELL_MANAGER_STATE.WAIT_TARGET)
				OR (eState = E_CELL_MANAGER_STATE.SELECT_FALLBACK)
				OR (eState = E_CELL_MANAGER_STATE.WAIT_MAGAZINE))))
		OR axMagazineExchangeInProgress[uiActiveMagazine]
		OR xUseAlternateMagazineForDetail
		OR xReselectMagazine)
	AND (NOT astMagazineStatus[uiActiveMagazine].xBusy
		OR axMagazineExchangeInProgress[uiActiveMagazine])
	AND NOT stRobotStatus.xBusy THEN
		IF xAlternateMagazineAvailable THEN
			IF uiActiveMagazine = UINT#1 THEN
				uiActiveMagazine := UINT#2;
			ELSE
				uiActiveMagazine := UINT#1;
			END_IF;
		ELSE
			// Без готовой замены старый код навечно оставлял магазин владельцем:
			// FB_MAGAZINE видел xRobotOwnsMagazine и не мог завершить Disable.
			// Освобождаем владение и ждём готовый магазин, не останавливая ячейку.
			uiActiveMagazine := UINT#0;
		END_IF;
		eMagazineOperation := E_MAGAZINE_OPERATION.NONE;
		eMachineOperation := E_MACHINE_OPERATION.NONE;
		uiSelectedMachine := UINT#0;
		uiSelectedType := UINT#0;
		iTakeSlot := SINT#0;
		iPutSlot := SINT#0;
		iTakeOriginSlot := SINT#0;
		IF uiActiveMagazine = UINT#0 THEN
			eState := E_CELL_MANAGER_STATE.WAIT_MAGAZINE;
		ELSE
			eState := E_CELL_MANAGER_STATE.PLAN_TARGET;
		END_IF;
	END_IF;
END_IF;

IF (uiActiveMagazine < UINT#1) OR (uiActiveMagazine > UINT#2) THEN
	IF uiPreferredMagazine > UINT#0 THEN
		uiActiveMagazine := uiPreferredMagazine;
	ELSIF xMagazine1Available THEN
		uiActiveMagazine := UINT#1;
	ELSIF xMagazine2Available THEN
		uiActiveMagazine := UINT#2;
	ELSE
		uiActiveMagazine := UINT#0;
	END_IF;
ELSIF NOT xRunning
AND (astMagazineStatus[uiActiveMagazine].xFinished
	OR astMagazineStatus[uiActiveMagazine].xError
	OR NOT astMagazineStatus[uiActiveMagazine].xEnabled
	OR xReselectMagazine) THEN
	IF (uiActiveMagazine <> UINT#1) AND xMagazine1Available THEN
		uiActiveMagazine := UINT#1;
	ELSIF (uiActiveMagazine <> UINT#2) AND xMagazine2Available THEN
		uiActiveMagazine := UINT#2;
	ELSIF xMagazine1Available THEN
		uiActiveMagazine := UINT#1;
	ELSIF xMagazine2Available THEN
		uiActiveMagazine := UINT#2;
	ELSE
		uiActiveMagazine := UINT#0;
	END_IF;
END_IF;

xActiveMagazineCanExchangeDetail := ((uiActiveMagazine = UINT#1) AND xMagazine1CanExchangeDetail)
	OR ((uiActiveMagazine = UINT#2) AND xMagazine2CanExchangeDetail);

IF (uiActiveMagazine >= UINT#1) AND (uiActiveMagazine <= UINT#2) THEN
	stMagazineStatus := astMagazineStatus[uiActiveMagazine];
	xActiveMagazineAutoSwapPending := axMagazineAutoSwapPending[uiActiveMagazine];
	xActiveMagazineExchangeInProgress := axMagazineExchangeInProgress[uiActiveMagazine];
ELSE
	stMagazineStatus := astMagazineStatus[1];
	xActiveMagazineAutoSwapPending := FALSE;
	xActiveMagazineExchangeInProgress := axMagazineExchangeInProgress[1];
END_IF;

// HOME_SAFETY — это диапазон вокруг именованной точки, а не требование
// побитового совпадения координат. Защёлка снимается только при принятом запуске:
// оператор не сможет подъехать к точке, снова отъехать и запустить цикл.
xRobotAtSafetyHome := (ABS(lrRobotActualX - stSafetyHomePoint.X) <= lrSafetyHomeToleranceX)
	AND (ABS(lrRobotActualY - stSafetyHomePoint.Y) <= lrSafetyHomeToleranceY)
	AND (ABS(lrRobotActualZ - stSafetyHomePoint.Z) <= lrSafetyHomeToleranceZ);

// Штатная остановка не требует HOME_SAFETY, пока робот остаётся в сохранённой
// позе. Любое последующее координатное перемещение (JOG, MoveAbsolute или
// MoveDirect) необратимо снимает доверие до следующего разрешённого запуска.
IF (eState = E_CELL_MANAGER_STATE.IDLE)
AND NOT xRunning
AND NOT xSafetyHomeRequired THEN
	IF NOT xStoppedPoseValid THEN
		lrStoppedPoseX := lrRobotActualX;
		lrStoppedPoseY := lrRobotActualY;
		lrStoppedPoseZ := lrRobotActualZ;
		xStoppedPoseValid := TRUE;
	ELSIF xManual
	AND ((ABS(lrRobotActualX - lrStoppedPoseX) > lrStoppedPoseTolerance)
	OR (ABS(lrRobotActualY - lrStoppedPoseY) > lrStoppedPoseTolerance)
	OR (ABS(lrRobotActualZ - lrStoppedPoseZ) > lrStoppedPoseTolerance)) THEN
		xSafetyHomeRequired := TRUE;
		xStoppedPoseValid := FALSE;
	END_IF;
END_IF;

// FB_ROBOT — источник фактического типа груза. Локальные значения менеджера
// принимаются от него после каждого цикла, что оставляет место для будущей
// инициализации зажатого захвата оператором.
IF stRobotStatus.xBlankAvailable THEN
	uiBlankPayloadType := stRobotStatus.uiBlankPayloadType;
ELSE
	uiBlankPayloadType := UINT#0;
END_IF;
IF stRobotStatus.xDetailAvailable THEN
	uiDetailPayloadType := stRobotStatus.uiDetailPayloadType;
ELSE
	uiDetailPayloadType := UINT#0;
END_IF;

// FB_MACHINE остаётся единственным владельцем таймаута запуска. Диспетчер только
// сохраняет короткое переходное состояние, чтобы новый цикл не исключался из прогноза.
FOR uiMachine := FIRST_MACHINE TO LAST_MACHINE DO
	IF axMachineStartPending[uiMachine]
	AND (astMachineStatus[uiMachine].xProcessing
		OR (astMachineStatus[uiMachine].ePartState = E_PART_STATE.EMPTY)
		OR NOT astMachineStatus[uiMachine].xEnabled
		OR astMachineStatus[uiMachine].xDisablePending
		OR astMachineStatus[uiMachine].xError) THEN
		axMachineStartPending[uiMachine] := FALSE;
	END_IF;
END_FOR;

Command.stRobot.xExecute := FALSE;
FOR uiGeometryIndex := UINT#1 TO UINT#2 DO
	GVL_GEOMETRY_CONTROL.astSignals[uiGeometryIndex].xReleased := FALSE;
END_FOR;
// После аварии контекст снимается лишь при подтверждённом выходе в HOME_SAFETY.
IF (uiGeometryStation >= UINT#1) AND (uiGeometryStation <= UINT#2)
AND (stRobotStatus.eCurrentPoint = E_POINT_NAME.HOME_SAFETY)
AND NOT stRobotStatus.xBusy AND NOT xMotionBusy
AND (eState <> E_CELL_MANAGER_STATE.GEOMETRY_DELIVER)
AND (eState <> E_CELL_MANAGER_STATE.GEOMETRY_RELEASE_COMMAND) THEN
	GVL_GEOMETRY_CONTROL.astSignals[uiGeometryStation].xReserve := FALSE;
	GVL_GEOMETRY_CONTROL.astSignals[uiGeometryStation].xDeposited := FALSE;
	GVL_GEOMETRY_CONTROL.astSignals[uiGeometryStation].xRobotInteraction := FALSE;
	GVL_GEOMETRY_CONTROL.astSignals[uiGeometryStation].xReleased := TRUE;
	IF xGeometryHeld AND (uiGeometryMachine >= UINT#1) AND (uiGeometryMachine <= UINT#3)
	AND stRobotStatus.xDetailAvailable THEN
		GVL_GEOMETRY_CONTROL.astCalls[uiGeometryMachine].uiStation := UINT#0;
		GVL_GEOMETRY_CONTROL.astCalls[uiGeometryMachine].uiState := UINT#2;
		GVL_GEOMETRY_CONTROL.astCalls[uiGeometryMachine].uiReason := UINT#4;
		F_GEOMETRY_EVENT(Call := GVL_GEOMETRY_CONTROL.astCalls[uiGeometryMachine]);
	END_IF;
	IF NOT stRobotStatus.xDetailAvailable THEN
		IF xGeometryHeld AND (uiGeometryMachine >= UINT#1) AND (uiGeometryMachine <= UINT#3) THEN
			IF (GVL_GEOMETRY_CONTROL.astCalls[uiGeometryMachine].uiState = UINT#2)
			OR (GVL_GEOMETRY_CONTROL.astCalls[uiGeometryMachine].uiState = UINT#3) THEN
				GVL_GEOMETRY_CONTROL.astCalls[uiGeometryMachine].uiState := UINT#7;
				GVL_GEOMETRY_CONTROL.astCalls[uiGeometryMachine].uiReason := UINT#5;
				F_GEOMETRY_EVENT(Call := GVL_GEOMETRY_CONTROL.astCalls[uiGeometryMachine]);
			END_IF;
		END_IF;
		xGeometryHeld := FALSE; uiGeometryMachine := UINT#0;
	END_IF;
	uiGeometryStation := UINT#0;
END_IF;
// Ручное изъятие из захвата после остановки завершает старый вызов. Подтверждённую
// укладку на ГК (state 4) этот путь не заменяет прерыванием и повторно не считает.
IF xGeometryHeld AND NOT stRobotStatus.xDetailAvailable AND NOT xRunning
AND NOT stRobotStatus.xBusy AND NOT xMotionBusy
AND (eState = E_CELL_MANAGER_STATE.IDLE)
AND (uiGeometryMachine >= UINT#1) AND (uiGeometryMachine <= UINT#3) THEN
	IF (GVL_GEOMETRY_CONTROL.astCalls[uiGeometryMachine].uiState = UINT#2)
	OR (GVL_GEOMETRY_CONTROL.astCalls[uiGeometryMachine].uiState = UINT#3) THEN
		GVL_GEOMETRY_CONTROL.astCalls[uiGeometryMachine].uiState := UINT#7;
		GVL_GEOMETRY_CONTROL.astCalls[uiGeometryMachine].uiReason := UINT#5;
		F_GEOMETRY_EVENT(Call := GVL_GEOMETRY_CONTROL.astCalls[uiGeometryMachine]);
	END_IF;
	xGeometryHeld := FALSE; uiGeometryMachine := UINT#0;
END_IF;
Command.stRobot.xStop := FALSE;
Command.stRobot.xReset := xReset;
Command.stRobot.eAction := E_ROBOT_ACTION.NONE;
Command.stRobot.eSetPoint := E_POINT_NAME.NONE;
Command.stRobot.iActiveSlot := SINT#0;
Command.stRobot.uiMagazineId := UINT#0;
Command.uiBlankPayloadType := uiBlankPayloadType;
Command.uiDetailPayloadType := uiDetailPayloadType;

Command.stMagazine.xEnable := FALSE;
Command.stMagazine.xDisable := FALSE;
Command.stMagazine.xExecute := FALSE;
Command.stMagazine.xStop := FALSE;
Command.stMagazine.eOperation := eMagazineOperation;
Command.stMagazine.iTakeSlot := iTakeSlot;
Command.stMagazine.iPutSlot := iPutSlot;
xChangePrepared := FALSE;

FOR uiMachine := FIRST_MACHINE TO LAST_MACHINE DO
	Command.axMachineExecute[uiMachine] := FALSE;
END_FOR;

uiReadyMachines := UINT#0;
xAnyMachineBusy := FALSE;
xMachineWorkPending := FALSE;
FOR uiMachine := FIRST_MACHINE TO LAST_MACHINE DO
	IF astMachineStatus[uiMachine].xBusy THEN
		xAnyMachineBusy := TRUE;
		xMachineWorkPending := TRUE;
	END_IF;
	IF astMachineStatus[uiMachine].xProcessing
	OR astMachineStatus[uiMachine].xPartReady
	OR axMachineStartPending[uiMachine]
	OR ((astMachineStatus[uiMachine].ePartState = E_PART_STATE.LOADED)
		AND ((astMachineStatus[uiMachine].ePartType = E_PART_TYPE.PART)
			OR (astMachineStatus[uiMachine].ePartType = E_PART_TYPE.DETAIL))) THEN
		xMachineWorkPending := TRUE;
	END_IF;
	IF IsMachineEligible(uiMachine := uiMachine) THEN
		uiReadyMachines := uiReadyMachines + UINT#1;
	END_IF;
END_FOR;

xRobotReady := NOT stRobotStatus.xBusy
	AND NOT stRobotStatus.xError;
xMagazineReady := (uiActiveMagazine >= UINT#1)
	AND (uiActiveMagazine <= UINT#2)
	AND NOT xActiveMagazineExchangeInProgress
	AND stMagazineStatus.xEnabled
	AND stMagazineStatus.xReady
	AND NOT stMagazineStatus.xBusy
	AND NOT stMagazineStatus.xError
	AND NOT stMagazineStatus.xFinished
	AND NOT stMagazineStatus.xDisablePending;

uiCandidateMachine := SelectMachineBeforeTake();
IF uiCandidateMachine = UINT#0 THEN
	uiCandidateMachine := SelectMachineForUnload(uiCurrentMachine := UINT#0);
END_IF;

// Для готовой детали пригоден только свободный слот её типа в магазине,
// который сейчас включён и доступен роботу. Свободная ячейка в отключённом
// или неисправном магазине не считается маршрутом.
xAnyMagazineDetailSlotAvailable := FALSE;
IF (uiDetailPayloadType >= UINT#1)
AND (uiDetailPayloadType <= Config.uiTypeCount) THEN
	FOR uiMagazineIndex := UINT#1 TO GVL_CELL_SETTINGS.MagazineCount DO
		IF astMagazineStatus[uiMagazineIndex].xEnabled
		AND astMagazineStatus[uiMagazineIndex].xReady
		AND NOT axMagazineExchangeInProgress[uiMagazineIndex]
		AND NOT astMagazineStatus[uiMagazineIndex].xBusy
		AND NOT astMagazineStatus[uiMagazineIndex].xError
		AND NOT astMagazineStatus[uiMagazineIndex].xFinished
		AND NOT astMagazineStatus[uiMagazineIndex].xDisablePending THEN
			IF astMagazineStatus[uiMagazineIndex].stTypeStatus.aiFreeSlot[uiDetailPayloadType] > SINT#0 THEN
				xAnyMagazineDetailSlotAvailable := TRUE;
			END_IF;
		END_IF;
	END_FOR;
END_IF;

// WARNING: место требуется только для готовой детали, уже находящейся у робота.
// Деталь в станке и полная палета заготовок при пустом роботе не создают W29.
// Взятие заготовки освобождает место; при двух грузах возможна загрузка станка.
// Штатный Stop снимает потребность в новом маршруте. Фронт проверяем отдельно:
// защёлка xStopRequested обновляется ниже, после регистрации предупреждений.
xNoDetailDestinationCondition := (xRunning OR rtStart.Q)
	AND NOT rtStop.Q
	AND NOT xStopRequested
	AND NOT xManual
	AND NOT xMagazineExchangeActive
	AND stRobotStatus.xDetailAvailable
	AND (uiDetailPayloadType >= UINT#1)
	AND (uiDetailPayloadType <= Config.uiTypeCount)
	AND NOT xAnyMagazineDetailSlotAvailable
	AND NOT xMagazine1CanExchangeDetail
	AND NOT xMagazine2CanExchangeDetail
	AND NOT xHeldBlankLoadAvailable
	AND ((eState = E_CELL_MANAGER_STATE.PLAN_TARGET)
		OR (eState = E_CELL_MANAGER_STATE.WAIT_TARGET)
		OR (eState = E_CELL_MANAGER_STATE.SELECT_FALLBACK)
		OR (eState = E_CELL_MANAGER_STATE.WAIT_MAGAZINE)
		OR (rtStart.Q AND (eState = E_CELL_MANAGER_STATE.IDLE)));

xNoBlankStockCondition := (xRunning OR rtStart.Q)
	AND NOT xManual
	AND NOT xMagazineExchangeActive
	AND NOT stRobotStatus.xBlankAvailable
	AND NOT stRobotStatus.xDetailAvailable
	AND astMagazineStatus[1].xOutBlank
	AND astMagazineStatus[2].xOutBlank
	AND NOT xMachineWorkPending
	AND (uiCandidateMachine = UINT#0)
	AND ((eState = E_CELL_MANAGER_STATE.PLAN_TARGET)
		OR (eState = E_CELL_MANAGER_STATE.WAIT_TARGET)
		OR (eState = E_CELL_MANAGER_STATE.WAIT_MAGAZINE)
		OR (rtStart.Q AND (eState = E_CELL_MANAGER_STATE.IDLE)));

CASE Config.uiTypeCount OF
	UINT#1: uiOperatorTypeMask := UINT#1;
	UINT#2: uiOperatorTypeMask := UINT#3;
	UINT#3: uiOperatorTypeMask := UINT#7;
ELSE
	uiOperatorTypeMask := UINT#0;
END_CASE;

// Для специального старта с двумя грузами оператор выбирает только среди действительно
// пустых, готовых и совместимых станков. Окончательная проверка выбора остаётся в PLC.
uiOperatorMachineMask := UINT#0;
IF (uiBlankPayloadType >= UINT#1)
AND (uiBlankPayloadType <= Config.uiTypeCount) THEN
	FOR uiMachine := FIRST_MACHINE TO LAST_MACHINE DO
		IF IsMachineCompatible(
			uiMachine := uiMachine,
			uiProductType := uiBlankPayloadType
		)
		AND astMachineStatus[uiMachine].xCanAcceptService
		AND (astMachineStatus[uiMachine].ePartState = E_PART_STATE.EMPTY) THEN
			CASE uiMachine OF
				UINT#1: uiOperatorMachineMask := uiOperatorMachineMask OR UINT#1;
				UINT#2: uiOperatorMachineMask := uiOperatorMachineMask OR UINT#2;
				UINT#3: uiOperatorMachineMask := uiOperatorMachineMask OR UINT#4;
			END_CASE;
		END_IF;
	END_FOR;
END_IF;

// Условия запуска публикуются раздельно: PLC остаётся единственным владельцем
// технологического решения, а HMI только объясняет его оператору.
xStartCheckCellIdle := (eState = E_CELL_MANAGER_STATE.IDLE) AND NOT xRunning;
xStartCheckAutomaticMode := NOT xManual;
xStartCheckNoBlockingError := NOT xGlobalError AND NOT xIoManual AND (Error.dwErrorActive = DWORD#0);
xStartCheckRobotInterfaceReady := xRobotInterfaceReady;
xStartCheckConfigurationValid := xConfigurationValid;
xStartCheckPointsConfigured := xPointsConfigured;
xStartCheckDrivesReady := xDrivesReady;
xStartCheckRobotReady := xRobotReady;
xStartCheckMagazineReady := xMagazineReady;
xStartCheckTaskAvailable := stRobotStatus.xBlankAvailable
		OR stRobotStatus.xDetailAvailable
		OR (uiCandidateMachine > UINT#0);
xStartCheckSafetyHome := NOT xSafetyHomeRequired OR xRobotAtSafetyHome;
xStartCheckSafety := xSafetyReady;

xReadyToStart := xStartCheckCellIdle
	AND xStartCheckAutomaticMode
	AND xStartCheckNoBlockingError
	AND xStartCheckRobotInterfaceReady
	AND xStartCheckConfigurationValid
	AND xStartCheckPointsConfigured
	AND xStartCheckDrivesReady
	AND xStartCheckRobotReady
	AND xStartCheckMagazineReady
	AND xStartCheckTaskAvailable
	AND xStartCheckSafetyHome
	AND xStartCheckSafety;

uiStartConditionsMet := UINT#0;
IF xStartCheckCellIdle THEN
	uiStartConditionsMet := uiStartConditionsMet + UINT#1;
END_IF;
IF xStartCheckAutomaticMode THEN
	uiStartConditionsMet := uiStartConditionsMet + UINT#1;
END_IF;
IF xStartCheckNoBlockingError THEN
	uiStartConditionsMet := uiStartConditionsMet + UINT#1;
END_IF;
IF xStartCheckRobotInterfaceReady THEN
	uiStartConditionsMet := uiStartConditionsMet + UINT#1;
END_IF;
IF xStartCheckConfigurationValid THEN
	uiStartConditionsMet := uiStartConditionsMet + UINT#1;
END_IF;
IF xStartCheckPointsConfigured THEN
	uiStartConditionsMet := uiStartConditionsMet + UINT#1;
END_IF;
IF xStartCheckDrivesReady THEN
	uiStartConditionsMet := uiStartConditionsMet + UINT#1;
END_IF;
IF xStartCheckRobotReady THEN
	uiStartConditionsMet := uiStartConditionsMet + UINT#1;
END_IF;
IF xStartCheckMagazineReady THEN
	uiStartConditionsMet := uiStartConditionsMet + UINT#1;
END_IF;
IF xStartCheckTaskAvailable THEN
	uiStartConditionsMet := uiStartConditionsMet + UINT#1;
END_IF;
IF xStartCheckSafetyHome THEN
	uiStartConditionsMet := uiStartConditionsMet + UINT#1;
END_IF;
IF xStartCheckSafety THEN
	uiStartConditionsMet := uiStartConditionsMet + UINT#1;
END_IF;

xFaultAllowed := (eState = E_CELL_MANAGER_STATE.IDLE)
	AND NOT xRunning
	AND NOT xGlobalError
	AND NOT xMotionBusy
	AND NOT stRobotStatus.xBusy
	AND NOT stMagazineStatus.xBusy
	AND NOT xAnyMachineBusy
	AND (Error.dwErrorActive = DWORD#0);
fbFaultInjector(Request := FaultRequest, xOwnerAllowed := xFaultAllowed);
FaultStatus := fbFaultInjector.Status;

IF fbFaultInjector.Status.xRejected THEN
	Diag.stWarning.uiCode := WRN_SIM_ERROR_NOT_ALLOWED;
	Diag.stWarning.udiSequence := Diag.stWarning.udiSequence + UDINT#1;
	IF Diag.stWarning.udiSequence = UDINT#0 THEN
		Diag.stWarning.udiSequence := UDINT#1;
	END_IF;
END_IF;

IF rtStart.Q
AND xSafetyHomeRequired
AND NOT xRobotAtSafetyHome
AND NOT (xRunning AND xStopRequested) THEN
	Diag.stWarning.uiCode := WRN_SAFETY_HOME_REQUIRED;
	Diag.stWarning.udiSequence := Diag.stWarning.udiSequence + UDINT#1;
	IF Diag.stWarning.udiSequence = UDINT#0 THEN
		Diag.stWarning.udiSequence := UDINT#1;
	END_IF;
ELSIF rtStart.Q AND NOT (xReadyToStart OR (xRunning AND xStopRequested)) THEN
	Diag.stWarning.uiCode := WRN_START_NOT_READY;
	Diag.stWarning.udiSequence := Diag.stWarning.udiSequence + UDINT#1;
	IF Diag.stWarning.udiSequence = UDINT#0 THEN
		Diag.stWarning.udiSequence := UDINT#1;
	END_IF;
END_IF;

IF rtStop.Q AND NOT xRunning THEN
	Diag.stWarning.uiCode := WRN_STOP_NOT_RUNNING;
	Diag.stWarning.udiSequence := Diag.stWarning.udiSequence + UDINT#1;
	IF Diag.stWarning.udiSequence = UDINT#0 THEN
		Diag.stWarning.udiSequence := UDINT#1;
	END_IF;
END_IF;

IF (uiModeRejectReason = UINT#2) OR (uiModeRejectReason = UINT#3) THEN
	IF uiModeRejectReason = UINT#2 THEN
		Diag.stWarning.uiCode := WRN_MANUAL_MODE_REJECTED;
	ELSE
		Diag.stWarning.uiCode := WRN_AUTOMATIC_MODE_REJECTED;
	END_IF;
	Diag.stWarning.udiSequence := Diag.stWarning.udiSequence + UDINT#1;
	IF Diag.stWarning.udiSequence = UDINT#0 THEN
		Diag.stWarning.udiSequence := UDINT#1;
	END_IF;
END_IF;

// Ответы HMI принимаются только пока PLC явно публикует активный шаг опроса.
xOperatorPromptState := (eState = E_CELL_MANAGER_STATE.WAIT_GRIPPER1_CONTENT)
	OR (eState = E_CELL_MANAGER_STATE.WAIT_GRIPPER1_TYPE)
	OR (eState = E_CELL_MANAGER_STATE.WAIT_GRIPPER2_CONTENT)
	OR (eState = E_CELL_MANAGER_STATE.WAIT_GRIPPER2_TYPE)
	OR (eState = E_CELL_MANAGER_STATE.WAIT_START_MACHINE);
xOperatorChoiceAllowed := xOperatorPromptState
	AND NOT xManual
	AND NOT xGlobalError
	AND (Error.dwErrorActive = DWORD#0)
	AND xRobotInterfaceReady
	AND xConfigurationValid
	AND xPointsConfigured
	AND xDrivesReady
	AND xRobotReady
	AND xMagazineReady
	AND (NOT xSafetyHomeRequired OR xRobotAtSafetyHome);
// Отмена не должна блокироваться из-за временно потерянной готовности:
// оператор всегда может закрыть незавершённый предпусковой опрос.
xOperatorCancelAllowed := xOperatorPromptState;

IF rtOperatorChoice.Q AND NOT xOperatorChoiceAllowed THEN
	Diag.stWarning.uiCode := WRN_OPERATOR_REPLY_REJECTED;
	Diag.stWarning.udiSequence := Diag.stWarning.udiSequence + UDINT#1;
	IF Diag.stWarning.udiSequence = UDINT#0 THEN
		Diag.stWarning.udiSequence := UDINT#1;
	END_IF;
END_IF;

IF rtOperatorCancel.Q THEN
	IF xOperatorCancelAllowed THEN
		uiBlankPayloadType := UINT#0;
		uiDetailPayloadType := UINT#0;
		uiSelectedMachine := UINT#0;
		uiSelectedType := UINT#0;
		eMachineOperation := E_MACHINE_OPERATION.NONE;
		eState := E_CELL_MANAGER_STATE.IDLE;
	ELSE
		Diag.stWarning.uiCode := WRN_OPERATOR_CANCEL_REJECTED;
		Diag.stWarning.udiSequence := Diag.stWarning.udiSequence + UDINT#1;
		IF Diag.stWarning.udiSequence = UDINT#0 THEN
			Diag.stWarning.udiSequence := UDINT#1;
		END_IF;
	END_IF;
END_IF;

// Если оператор или внешний контроллер изменил захваты во время вопроса, старый ответ больше недостоверен.
IF xOperatorPromptState
AND NOT rtOperatorCancel.Q
AND ((stRobotStatus.xBlankAvailable <> xPrestartGripper1Occupied)
	OR (stRobotStatus.xDetailAvailable <> xPrestartGripper2Occupied)) THEN
	Diag.stWarning.uiCode := WRN_OPERATOR_REPLY_REJECTED;
	Diag.stWarning.udiSequence := Diag.stWarning.udiSequence + UDINT#1;
	IF Diag.stWarning.udiSequence = UDINT#0 THEN
		Diag.stWarning.udiSequence := UDINT#1;
	END_IF;
	uiBlankPayloadType := UINT#0;
	uiDetailPayloadType := UINT#0;
	eState := E_CELL_MANAGER_STATE.IDLE;
END_IF;

IF xOperatorPromptState
AND xManual THEN
	uiBlankPayloadType := UINT#0;
	uiDetailPayloadType := UINT#0;
	uiSelectedMachine := UINT#0;
	uiSelectedType := UINT#0;
	eMachineOperation := E_MACHINE_OPERATION.NONE;
	eState := E_CELL_MANAGER_STATE.IDLE;
END_IF;

// Условия ожидания не являются ошибкой и не останавливают ячейку. Каждое
// предупреждение регистрируется один раз на непрерывный эпизод; после очистки
// причины новое появление условия создаст новую запись журнала.
IF xNoDetailDestinationCondition
AND NOT xDetailDestinationWarningActive THEN
	Diag.stWarning.uiCode := WRN_NO_DETAIL_DESTINATION;
	Diag.stWarning.udiSequence := Diag.stWarning.udiSequence + UDINT#1;
	IF Diag.stWarning.udiSequence = UDINT#0 THEN
		Diag.stWarning.udiSequence := UDINT#1;
	END_IF;
END_IF;
xDetailDestinationWarningActive := xNoDetailDestinationCondition;

IF xNoBlankStockCondition
AND NOT xBlankStockWarningActive THEN
	Diag.stWarning.uiCode := WRN_NO_BLANK_STOCK;
	Diag.stWarning.udiSequence := Diag.stWarning.udiSequence + UDINT#1;
	IF Diag.stWarning.udiSequence = UDINT#0 THEN
		Diag.stWarning.udiSequence := UDINT#1;
	END_IF;
END_IF;
xBlankStockWarningActive := xNoBlankStockCondition;

IF rtStop.Q OR xManual THEN
	xStopRequested := TRUE;
ELSIF rtStart.Q AND xRunning
AND (eState <> E_CELL_MANAGER_STATE.MACHINE_FAULT_STOP) THEN
	xStopRequested := FALSE;
END_IF;

// Ошибка робота становится ошибкой автоматического цикла только когда ячейка
// действительно выполняет цикл. В IDLE ручная ошибка остаётся у своего
// первичного владельца (ось, группа или робот) и не создаёт ложный каскад.
IF xRunning AND stRobotStatus.xError THEN
	xSafetyHomeRequired := TRUE;
	xStoppedPoseValid := FALSE;
	Error.dwErrorActive := Error.dwErrorActive OR ERR_ROBOT;
	eState := E_CELL_MANAGER_STATE.ERROR;
END_IF;

IF xGlobalError
AND (eState <> E_CELL_MANAGER_STATE.IDLE)
AND (eState <> E_CELL_MANAGER_STATE.ERROR) THEN
	// Не каждая общая авария требует возврата. Защёлкиваем только ситуацию,
	// где прервано движение либо робот мог находиться внутри станка/магазина.
	IF stRobotStatus.xBusy
	OR xMotionBusy
	OR (eState = E_CELL_MANAGER_STATE.ROUTE_TO_TARGET)
	OR (eState = E_CELL_MANAGER_STATE.RELEASE_ROBOT_COMMAND)
	OR (eState = E_CELL_MANAGER_STATE.SERVICE_TARGET)
	OR (eState = E_CELL_MANAGER_STATE.MAGAZINE_EXECUTE)
	OR (eState = E_CELL_MANAGER_STATE.RELEASE_MAGAZINE)
	OR (eState = E_CELL_MANAGER_STATE.MACHINE_FAULT_STOP) THEN
		xSafetyHomeRequired := TRUE;
		xStoppedPoseValid := FALSE;
	END_IF;
	Error.dwErrorActive := Error.dwErrorActive OR ERR_GLOBAL_STOP;
	eState := E_CELL_MANAGER_STATE.ERROR;
END_IF;

// Штатный Stop ждёт безопасную технологическую границу. Тестовый Abort ждать
// её не должен: удерживаем Stop владельцев и не даём автоматам выдать новую
// команду, пока Motion фактически не закончил торможение.
IF xTestAbort THEN
	eState := E_CELL_MANAGER_STATE.TEST_ABORT_STOP;
END_IF;

// При передаче I/O оператору нельзя ждать программные Busy: именно зависший
// владелец может требовать восстановления. Аварии и физический груз сохраняются.
IF xIoManual THEN
	xRunning := FALSE;
	xStopRequested := FALSE;
	xMachineServiceStarted := FALSE;
	xReselectAfterRobotRelease := FALSE;
	xSafetyHomeRequired := TRUE;
	xStoppedPoseValid := FALSE;
	uiSelectedMachine := UINT#0;
	uiSelectedType := UINT#0;
	eMachineOperation := E_MACHINE_OPERATION.NONE;
	eMagazineOperation := E_MAGAZINE_OPERATION.NONE;
	iTakeSlot := SINT#0;
	iPutSlot := SINT#0;
	iTakeOriginSlot := SINT#0;
	FOR uiMachine := FIRST_MACHINE TO LAST_MACHINE DO
		axMachineStartPending[uiMachine] := FALSE;
	END_FOR;
	IF eState <> E_CELL_MANAGER_STATE.ERROR THEN
		eState := E_CELL_MANAGER_STATE.IDLE;
	END_IF;
END_IF;

// ГК не зависит от готовности палет. Если магазин потерян после выгрузки,
// сначала доставляем вызванную деталь на свободный ГК либо паркуемся у занятого.
IF xRunning AND xGeometryHeld AND stRobotStatus.xDetailAvailable
AND (eState = E_CELL_MANAGER_STATE.WAIT_MAGAZINE)
AND NOT stRobotStatus.xBusy AND NOT xMotionBusy THEN
	PlanGeometry();
END_IF;

CASE eState OF
	E_CELL_MANAGER_STATE.IDLE:
		xRunning := FALSE;
		xStopRequested := FALSE;
		xMachineServiceStarted := FALSE;
		xReselectAfterRobotRelease := FALSE;
		eMagazineOperation := E_MAGAZINE_OPERATION.NONE;
		IF fbFaultInjector.xBothGrippers THEN
			Error.dwErrorActive := Error.dwErrorActive OR ERR_BOTH_GRIPPERS;
			eState := E_CELL_MANAGER_STATE.ERROR;
		ELSIF rtStart.Q AND NOT xManual THEN
			IF xReadyToStart THEN
				xPrestartGripper1Occupied := stRobotStatus.xBlankAvailable;
				xPrestartGripper2Occupied := stRobotStatus.xDetailAvailable;
				uiBlankPayloadType := UINT#0;
				uiDetailPayloadType := UINT#0;
				uiSelectedMachine := UINT#0;
				uiSelectedType := UINT#0;
				eMachineOperation := E_MACHINE_OPERATION.NONE;
				// Новый Start заново идентифицирует уже находящийся в захвате груз.
				// Слот происхождения прошлого цикла к нему не относится: иначе
				// RETURN_BLANK может попытаться положить груз в занятый чужой слот.
				iTakeSlot := SINT#0;
				iPutSlot := SINT#0;
				iTakeOriginSlot := SINT#0;
				eState := E_CELL_MANAGER_STATE.PRESTART_IDENTIFY;
			END_IF;
		END_IF;

	E_CELL_MANAGER_STATE.PRESTART_IDENTIFY:
		IF xManual THEN
			eState := E_CELL_MANAGER_STATE.IDLE;
		ELSIF xPrestartGripper1Occupied THEN
			eState := E_CELL_MANAGER_STATE.WAIT_GRIPPER1_CONTENT;
		ELSIF xPrestartGripper2Occupied THEN
			eState := E_CELL_MANAGER_STATE.WAIT_GRIPPER2_CONTENT;
		ELSE
			xSafetyHomeRequired := FALSE;
			xStoppedPoseValid := FALSE;
			xRunning := TRUE;
			eState := E_CELL_MANAGER_STATE.PLAN_TARGET;
		END_IF;

